(* IEC 61131-3 sources: daoli-st-library/DL_Process (part 52) *)

(* ---- FB_DL_SputterTargetBurnInSeq.st ---- *)
//==============================================================================
// 功能块：FB_DL_SputterTargetBurnInSeq ｜ 中文名称：溅射靶预烧与功率爬坡序（复杂度 C4）
// 所属子库：DL_Process ｜ 版本 VERSION: v1.0.0 ｜ 兼容：CODESYS V3.5+ / TwinCAT 3 / 汇川 InoProShop
// 功能描述：新靶装机后的预烧处理——真空达标 → 通 Ar 稳气 → 功率按斜率爬升 → 预烧到规定
//           能量 → 按斜率降功率 → 关快门 → 关气 → 完成。全程统计打火次数，超限立即把功率
//           指令压到 0 并锁存 xArcTrip；中止与打火停机一律走三段关断序（降功率 → 关快门
//           → 关气），禁单拍全断（会污染靶面）。
// 开源溯源 (Origin)：道莅原创实现（参考 SEMI F47 与磁控溅射靶预烧工艺惯例 分类与参数
//           域，许可证=MIT，借鉴点=「按斜率爬升 + 累计能量达量停烧 + 打火计数联锁」的
//           预烧序）
// 单位表：气压[Pa] / 功率[kW] / 能量[kWh] / 斜率[kW/s] / 打火[次] / 时间[ms]
// 能量离散积分（本件核心积分，换算写清）：
//   fEnergyKWh = Σ (P[kW] × Δt[s]) ÷ 3600 [s/h]；由 W 折算 kW 的 ÷1000 已含在入口量纲
//   上（若上层以 W 给功率，须先 ÷1000 再进本件），Δt 取 DL_SPT_DT_S 假定 10 ms 周期。
// 错误码表（Process 段 0005，故障窗口 3F11~3F19，信息窗口 3F91）：
//   16#0005_3F11 故障级：组态非法（设定压/容差/设定功率/斜率/能量 <= 0 或打火上限 = 0）
//   16#0005_3F12 故障级：实时量入口非有限（腔压 / 功率 NaN 或 Inf）或幅值超上限，拒算
//   16#0005_3F13 故障级：真空未达标超时（tRampTimeout 内气压未进入设定带）
//   16#0005_3F14 故障级：稳气超时（tRampTimeout 内气压未在带内稳住 tGasStabTime）
//   16#0005_3F15 故障级：功率爬坡超时（tRampTimeout 内未爬到设定功率）
//   16#0005_3F16 故障级：预烧超时（tBurnTimeout 内累计能量未达 fBurnEnergyKWh）
//   16#0005_3F17 故障级：打火超限（累计打火 > nArcLimit，功率立即压 0 并锁存 xArcTrip）
//   16#0005_3F18 故障级：关断序超时（降功率/关快门/关气任一段超 tRampTimeout）
//   16#0005_3F19 故障级兜底：状态机落 ELSE 非法态，全输出断
//   16#0005_3F91 信息级：预烧完成（进入 eDone 拍，不置 bError）
//           故障级码全部锁存回放（R187），唯一清除路径 = bReset 上升沿（含打火锁存）。
// 状态机：E_DL_SputterBurnState（八态：eIdle=0 / eVacCheck=10 / eGasStab=20 / eRampUp=30 /
//           eBurnIn=40 / eRampDown=50 / eDone=60 / eFault=99）。三段关断序不占相位，由
//           内部段号 _uDownStage 驱动（0 降功率 / 1 关快门 / 2 关气）。
// 边界行为：① 真空或气压未进带绝不加功率（eRampUp 入口以 _bVacOk 为唯一前提）；② 打火
//           超限属最高优先级：段 5 在功率生成处先判 _bArcTrip 并压 0，不等状态机；③ 三段
//           关断序每段之间留物理动作时间（DL_SPT_SHUTTER_T / DL_SPT_GAS_T），禁单拍全断；
//           ④ 中止与打火停机共用同一关断序，关断后落 eFault 或 eDone 由 _bArcTrip 决定；
//           ⑤ 八态 CASE 每态显式 + ELSE 兜底 → 3F19 全断。
// 语义假设：① nArcCount 为打火探测器累计计数，本件按增量累加并对上游复位做单调化处理；
//           ② 快门开 = xShutterCmd TRUE 表示靶面暴露给基片，预烧期按工艺允许开快门（挡板
//           由上层另控）；③ 腔压判据用绝对偏差带，不含符号方向。
// 依赖纪律：仅 Standard.library（TON / R_TRIG）；零 GVL、零 VAR_EXTERNAL、零物理地址。
// 修订历史：v1.0.0 2026-11-25 R88 首版（无人值守批次 · 复杂件 C4 · 序号 4）
//==============================================================================

(*------------------------------------------------------------------------------
 * 枚举: E_DL_SputterBurnState（归属本功能块，同文件发布，全库唯一定义）
 * 含义: 预烧相位，与段 8 状态机、段 9 输出置位一一对应。
 *-----------------------------------------------------------------------------*)
TYPE E_DL_SputterBurnState :
(
    eIdle     := 0,  // 空闲：等启动沿 / Idle, awaiting the start edge
    eVacCheck := 10, // 真空核对：腔压进入设定带 / Vacuum check against the pressure band
    eGasStab  := 20, // 稳气：通 Ar 并在带内稳住规定时间 / Argon stabilisation inside the band
    eRampUp   := 30, // 功率爬坡：按斜率爬到设定功率 / Power ramp up to the setpoint
    eBurnIn   := 40, // 预烧：累计能量到量前持续 / Burn-in until the energy target is met
    eRampDown := 50, // 降功率与三段关断 / Power ramp down and the three-stage shutdown
    eDone     := 60, // 完成：预烧结束 / Done, burn-in finished
    eFault    := 99  // 故障：组态/超时/打火/非法态 / Fault, configuration, timeout, arcing or illegal state
);
END_TYPE

FUNCTION_BLOCK FB_DL_SputterTargetBurnInSeq
VAR_INPUT
    xEnable       : BOOL;   // 使能，FALSE 期间按中止处理（走三段关断） [—] / Enable, a drop aborts into the shutdown
    xStart        : BOOL;   // 启动请求，上升沿生效 [—] / Start request, rising edge effective
    xAbort        : BOOL;   // 中止请求，任意拍生效（走三段关断） [—] / Abort request, moves into the shutdown
    xReset        : BOOL;   // 故障复位，上升沿清全部锁存（含打火锁存） [—] / Fault reset, clears all latches
    fChamberPressPa : LREAL; // 腔体实际气压 [Pa] / Actual chamber pressure [Pa]
    fPressSetPa   : LREAL;  // 工艺设定气压 [Pa]，须 > 0 / Process pressure setpoint [Pa]
    fPressTolPa   : LREAL;  // 气压允许偏差 [Pa]，须 > 0 / Allowed pressure tolerance [Pa]
    fPowerKW      : LREAL;  // 实际输出功率 [kW] / Actual delivered power [kW]
    fPowerSetKW   : LREAL;  // 预烧设定功率 [kW]，须 > 0 / Burn-in power setpoint [kW]
    fRampKWperS   : LREAL;  // 功率爬坡/降坡斜率 [kW/s]，须 > 0 / Power ramp rate [kW/s]
    fBurnEnergyKWh: LREAL;  // 预烧目标能量 [kWh]，须 > 0 / Burn-in energy target [kWh]
    nArcCount     : UDINT;  // 打火探测器累计计数 [次] / Arc detector accumulated count
    nArcLimit     : UDINT;  // 打火累计上限 [次]，须 > 0 / Accumulated arc ceiling
    tGasStabTime  : TIME;   // 稳气时长 [ms] / Gas stabilisation time [ms]
    tRampTimeout  : TIME;   // 真空/稳气/爬坡/关断超时 [ms] / Vacuum, gas, ramp and shutdown timeout [ms]
    tBurnTimeout  : TIME;   // 预烧最长允许时间 [ms] / Maximum burn-in time [ms]
END_VAR
VAR_OUTPUT
    fPowerCmdKW     : LREAL;  // 功率指令出口 [kW]，0 = 断功率 / Power command outlet [kW], 0 = off
    xArValveCmd     : BOOL;   // 氩气进气阀命令 [—] / Argon inlet valve command
    xShutterCmd     : BOOL;   // 快门命令（TRUE = 开） [—] / Shutter command, TRUE = open
    bRunning        : BOOL;   // 预烧进行中（非空闲非完成非故障） [—] / Burn-in active
    bDone           : BOOL;   // 预烧完成相电平 [—] / Burn-in done, level in the done phase
    bError          : BOOL;   // 故障级标志，仅故障级码置位 [—] / Fault-class flag, fault-level codes only
    nErrCode        : UDINT;  // 错误码，0 = 无错 [—] / Error code, 0 = none
    fEnergyKWh      : LREAL;  // 累计预烧能量 [kWh] / Accumulated burn-in energy [kWh]
    nArcTotal       : UDINT;  // 累计打火次数 [次] / Accumulated arc count
    xArcTrip        : BOOL;   // 打火超限锁存（bReset 清） [—] / Arc trip latch, cleared by bReset
END_VAR
VAR
    _eState         : E_DL_SputterBurnState := E_DL_SputterBurnState.eIdle; // 当前相位 [—] / Current phase
    _bInit          : BOOL := FALSE;  // 首扫标志，取非判定 [—] / First-scan flag, tested negated
    _fPowerCmd      : LREAL;          // 功率指令斜率限幅后的保持量 [kW] / Held command after rate limiting [kW]
    _fEnergyKWh     : LREAL;          // 内部累计能量 [kWh] / Internal accumulated energy [kWh]
    _nArcTotal      : UDINT;          // 内部累计打火次数 [次] / Internal accumulated arc count
    _nArcPrev       : UDINT;          // 上拍打火计数快照 [次] / Previous-scan arc count snapshot
    _bCfgBad        : BOOL;           // 组态非法锁存 / Illegal configuration latch
    _bCfgOk         : BOOL;           // 本拍组态合法（派生量不锁存） [—] / Configuration legal this scan
    _bSigBad        : BOOL;           // 实时量非有限锁存 / Non-finite process value latch
    _bVacOk         : BOOL;           // 气压在设定带内（派生量） [—] / Pressure inside the setpoint band
    _bArcTrip       : BOOL;           // 打火超限锁存 / Arc trip latch
    _bVacTmo        : BOOL;           // 真空超时锁存 / Vacuum timeout latch
    _bGasTmo        : BOOL;           // 稳气超时锁存 / Gas stabilisation timeout latch
    _bRampTmo       : BOOL;           // 爬坡超时锁存 / Ramp timeout latch
    _bBurnTmo       : BOOL;           // 预烧超时锁存 / Burn-in timeout latch
    _bDownTmo       : BOOL;           // 关断序超时锁存 / Shutdown timeout latch
    _bIllegal       : BOOL;           // 非法状态标志 / Illegal state flag
    _bInfoDone      : BOOL;           // 预烧完成信息当拍标志 / Burn-in done info flag of this scan
    _bAbortReq      : BOOL;           // 中止请求合成（xAbort 或失能） [—] / Combined abort request
    _uDownStage     : UINT;           // 关断段号 0=降功率 1=关快门 2=关气 / Shutdown stage 0 power 1 shutter 2 gas
    rtStart         : R_TRIG;         // 启动沿，段 7 无条件刷新 [—] / Start edge, refreshed in segment 7
    rtReset         : R_TRIG;         // 复位沿，段 7 无条件刷新 [—] / Reset edge, refreshed in segment 7
    tonVac          : TON;            // 真空核对超时 [ms] / Vacuum check timeout [ms]
    tonGas          : TON;            // 稳气计时（仅在带内累计） [ms] / Gas stabilisation timer inside the band
    tonGasMax       : TON;            // 稳气最长允许时间 [ms] / Maximum stabilisation time [ms]
    tonRamp         : TON;            // 功率爬坡超时 [ms] / Ramp timeout [ms]
    tonBurn         : TON;            // 预烧最长允许时间 [ms] / Maximum burn-in time [ms]
    tonShutter      : TON;            // 关快门动作让位 [ms] / Shutter travel dwell [ms]
    tonGasClose     : TON;            // 关气动作让位 [ms] / Gas closing dwell [ms]
    tonDownMax      : TON;            // 关断序总超时 [ms] / Total shutdown timeout [ms]
END_VAR
VAR CONSTANT
    DL_EPS           : LREAL := 1.0E-9;      // 浮点容差零点，兼作除法分母下限 / Float epsilon, also the divisor floor
    DL_SPT_DT_S      : LREAL := 0.01;        // 爬坡与积分的假定任务周期 [s]（10 ms） / Assumed task period [s]
    DL_SPT_SEC_PER_H : LREAL := 3600.0;      // 秒折算小时 [s/h]，能量积分用 / Seconds per hour for the energy integral
    DL_SPT_POW_EPS   : LREAL := 0.05;        // 功率到位容差 [kW] / Power arrival tolerance [kW]
    DL_SPT_POWER_MAX : LREAL := 500.0;       // 功率反馈合法幅值上限 [kW] / Legal power ceiling [kW]
    DL_SPT_PRESS_MAX : LREAL := 100000.0;    // 气压反馈合法幅值上限 [Pa] / Legal pressure ceiling [Pa]
    DL_SPT_SHUTTER_T : TIME  := T#800MS;     // 关快门动作让位 [ms] / Shutter travel dwell [ms]
    DL_SPT_GAS_T     : TIME  := T#500MS;     // 关气动作让位 [ms] / Gas closing dwell [ms]
END_VAR
(*------------------------------------------------------------------------------
 * 段 1｜每拍预置：全部输出先落安全侧，单拍标志预清零
 *      All outputs preset to the safe side, one-shot flags pre-cleared
 *-----------------------------------------------------------------------------*)
fPowerCmdKW := 0.0;                         // 功率指令先归零（安全侧） / Power command zeroed first
xArValveCmd := FALSE; xShutterCmd := FALSE; // 氩气与快门命令先断 / Argon and shutter commands cleared
bRunning := FALSE;  bDone := FALSE;         // 运行与完成标志每拍重算 / Running and done flags recomputed
bError := FALSE;    nErrCode := 16#0000_0000; // 故障标志与错误码每拍重算 / Fault flag and code recomputed
_bIllegal := FALSE; _bInfoDone := FALSE;    // 非法态与完成信息预清零 / Illegal and done-info flags pre-cleared

(*------------------------------------------------------------------------------
 * 段 2｜首扫初始化：相位、指令保持量、能量、打火累计与关断段号复位
 *      First-scan initialisation of phase, command, energy, arc count and stage
 *-----------------------------------------------------------------------------*)
IF NOT _bInit THEN
    _eState     := E_DL_SputterBurnState.eIdle; // 相位从空闲起步 / Phase starts idle
    _fPowerCmd := 0.0;  _fEnergyKWh := 0.0;     // 指令与能量从零起步 / Command and energy start at zero
    _nArcTotal := 0;    _nArcPrev  := 0;  _uDownStage := 0; // 打火累计/快照/关断段号从零起步 / Arc, snapshot and stage zero
    _bInit := TRUE;                             // 首扫只做一次 / The first scan runs once
END_IF
(*------------------------------------------------------------------------------
 * 段 3｜实时量入口非有限闸 + 组态闸 + 气压带判据
 *      Non-finite inlet gate, configuration gates and the pressure band criterion
 *-----------------------------------------------------------------------------*)
IF NOT (fChamberPressPa > -1.0E30 AND fChamberPressPa < 1.0E30) THEN _bSigBad := TRUE; END_IF  // 腔压非有限 → 3F12 / Non-finite pressure, 3F12
IF ABS(fChamberPressPa) > DL_SPT_PRESS_MAX THEN _bSigBad := TRUE; END_IF                     // 腔压幅值超上限 → 3F12 / Beyond the ceiling, 3F12
IF NOT (fPowerKW > -1.0E30 AND fPowerKW < 1.0E30) THEN _bSigBad := TRUE; END_IF               // 功率非有限 → 3F12 / Non-finite power, 3F12
IF ABS(fPowerKW) > DL_SPT_POWER_MAX THEN _bSigBad := TRUE; END_IF                             // 功率幅值超上限 → 3F12 / Beyond the ceiling, 3F12
IF NOT (fPressSetPa > -1.0E30 AND fPressSetPa < 1.0E30) THEN _bCfgBad := TRUE; END_IF         // 设定压非有限 → 3F11 / Non-finite setpoint pressure, 3F11
IF NOT (fPowerSetKW > -1.0E30 AND fPowerSetKW < 1.0E30) THEN _bCfgBad := TRUE; END_IF         // 设定功率非有限 → 3F11 / Non-finite setpoint power, 3F11
IF NOT (fRampKWperS > -1.0E30 AND fRampKWperS < 1.0E30) THEN _bCfgBad := TRUE; END_IF         // 斜率非有限 → 3F11 / Non-finite ramp, 3F11
IF NOT (fBurnEnergyKWh > -1.0E30 AND fBurnEnergyKWh < 1.0E30) THEN _bCfgBad := TRUE; END_IF    // 目标能量非有限 → 3F11 / Non-finite energy, 3F11
IF (fPressSetPa <= DL_EPS) OR (fPressTolPa <= DL_EPS) OR (fPowerSetKW <= DL_EPS)
   OR (fRampKWperS <= DL_EPS) OR (fBurnEnergyKWh <= DL_EPS) THEN _bCfgBad := TRUE; END_IF // 五者须为正 → 3F11 / All five must be positive
IF nArcLimit = 0 THEN _bCfgBad := TRUE; END_IF                          // 打火上限为 0 即永久跳闸 → 3F11 / Zero arc limit, 3F11
IF (tGasStabTime <= T#0MS) OR (tRampTimeout <= T#0MS) OR (tBurnTimeout <= T#0MS) THEN _bCfgBad := TRUE; END_IF // 时间量须为正 → 3F11
_bCfgOk := NOT _bCfgBad;                    // 本拍组态合法派生量 / Configuration-legal derived flag of this scan
_bVacOk := ABS(fChamberPressPa - fPressSetPa) <= fPressTolPa; // 气压带判据 [Pa] / Pressure band criterion [Pa]

(*------------------------------------------------------------------------------
 * 段 4｜打火累计（增量单调化）与超限锁存
 *      Arc accumulation with monotonic handling of an upstream counter reset
 *-----------------------------------------------------------------------------*)
IF nArcCount >= _nArcPrev THEN _nArcTotal := _nArcTotal + (nArcCount - _nArcPrev); // 增量累加 / Increment accumulated
ELSE _nArcTotal := _nArcTotal + nArcCount; END_IF                                  // 上游复位按新窗累加 / Upstream reset, new window
_nArcPrev := nArcCount;                     // 计数快照推进 / Count snapshot advanced
IF (_nArcTotal > nArcLimit) THEN
    _bArcTrip := TRUE;                      // 打火超限锁存 → 3F17 / Arc ceiling exceeded, 3F17
END_IF

(*------------------------------------------------------------------------------
 * 段 5｜功率指令生成（打火优先压 0）+ 斜率限幅 + 能量离散积分
 *      Power command generation, arc-first zeroing, rate limiting and energy integral
 *-----------------------------------------------------------------------------*)
IF _bArcTrip THEN
    _fPowerCmd := 0.0;                      // 打火超限：功率立即压 0（不等状态机） / Arc trip, power forced to zero
ELSIF (_eState = E_DL_SputterBurnState.eRampUp) OR (_eState = E_DL_SputterBurnState.eBurnIn) THEN
    IF fPowerSetKW > _fPowerCmd THEN
        _fPowerCmd := _fPowerCmd + fRampKWperS * DL_SPT_DT_S;       // 升坡 [kW] / Ramp up [kW]
        IF _fPowerCmd > fPowerSetKW THEN _fPowerCmd := fPowerSetKW; END_IF // 上钳设定值 / Clamp at setpoint
    ELSIF fPowerSetKW < _fPowerCmd THEN
        _fPowerCmd := _fPowerCmd - fRampKWperS * DL_SPT_DT_S;       // 降坡 [kW] / Ramp down [kW]
        IF _fPowerCmd < fPowerSetKW THEN _fPowerCmd := fPowerSetKW; END_IF // 下钳设定值 / Clamp at setpoint
    END_IF
ELSIF _eState = E_DL_SputterBurnState.eRampDown THEN
    _fPowerCmd := _fPowerCmd - fRampKWperS * DL_SPT_DT_S;           // 关断序段 0：降功率 [kW] / Shutdown stage 0, ramp down
    IF _fPowerCmd < 0.0 THEN _fPowerCmd := 0.0; END_IF              // 下钳 0 / Lower clamp at zero
ELSE
    _fPowerCmd := 0.0;                      // 其余相指令归零 / Zeroed in all other phases
END_IF
IF (_eState = E_DL_SputterBurnState.eBurnIn) AND (DL_SPT_SEC_PER_H > DL_EPS) THEN
    _fEnergyKWh := _fEnergyKWh + (_fPowerCmd * DL_SPT_DT_S) / DL_SPT_SEC_PER_H; // 能量积分 [kWh] / Energy integral [kWh]
END_IF
fPowerCmdKW := _fPowerCmd; fEnergyKWh := _fEnergyKWh; // 功率指令与能量出口 [kW]/[kWh] / Power and energy outlets
nArcTotal := _nArcTotal;    xArcTrip := _bArcTrip;    // 累计打火与打火锁存出口 / Arc count and arc trip outlets

(*------------------------------------------------------------------------------
 * 段 6｜中止入口（任意运行相 → 三段关断序）与复位
 *      Abort entry into the three-stage shutdown plus the reset edge
 *-----------------------------------------------------------------------------*)
_bAbortReq := xAbort OR (NOT xEnable);      // 中止请求合成：显式中止或失能 / Combined abort: explicit abort or enable loss
IF _bAbortReq AND (_eState <> E_DL_SputterBurnState.eIdle) AND (_eState <> E_DL_SputterBurnState.eRampDown)
   AND (_eState <> E_DL_SputterBurnState.eDone) AND (_eState <> E_DL_SputterBurnState.eFault) THEN
    _uDownStage := 0;                       // 关断序从段 0（降功率）起 / Shutdown starts at stage 0
    _eState     := E_DL_SputterBurnState.eRampDown; // 进关断相 / To the shutdown phase
END_IF
IF rtReset.Q THEN
    _bCfgBad := FALSE;  _bSigBad := FALSE;  _bArcTrip := FALSE; // 复位清组态/入口/打火锁存 / Clears configuration, inlet and arc latches
    _bVacTmo := FALSE;  _bGasTmo := FALSE;  _bRampTmo := FALSE; // 复位清真空/稳气/爬坡锁存 / Clears vacuum, gas and ramp latches
    _bBurnTmo := FALSE; _bDownTmo := FALSE;                     // 复位清预烧/关断锁存 / Clears burn-in and shutdown latches
END_IF
(*------------------------------------------------------------------------------
 * 段 7｜定时器与边沿无条件周期刷新（R7：CASE 之外每拍必调，各司其职不复用）
 *      Timers and edges refreshed unconditionally every scan, outside the CASE
 *-----------------------------------------------------------------------------*)
rtStart(CLK := xStart); rtReset(CLK := xReset); // 启动沿与复位沿无条件刷新 / Start and reset edges refreshed
tonVac(IN := (_eState = E_DL_SputterBurnState.eVacCheck), PT := tRampTimeout);                     // 真空核对超时 / Vacuum timeout
tonGas(IN := (_eState = E_DL_SputterBurnState.eGasStab) AND _bVacOk, PT := tGasStabTime);          // 带内稳气计时 / In-band gas timer
tonGasMax(IN := (_eState = E_DL_SputterBurnState.eGasStab), PT := tRampTimeout);                   // 稳气最长允许 / Maximum stabilisation
tonRamp(IN := (_eState = E_DL_SputterBurnState.eRampUp), PT := tRampTimeout);                      // 爬坡超时 / Ramp timeout
tonBurn(IN := (_eState = E_DL_SputterBurnState.eBurnIn), PT := tBurnTimeout);                      // 预烧超时 / Burn-in timeout
tonShutter(IN := (_eState = E_DL_SputterBurnState.eRampDown) AND (_uDownStage = 1), PT := DL_SPT_SHUTTER_T); // 关快门让位 / Shutter dwell
tonGasClose(IN := (_eState = E_DL_SputterBurnState.eRampDown) AND (_uDownStage = 2), PT := DL_SPT_GAS_T);    // 关气让位 / Gas dwell
tonDownMax(IN := (_eState = E_DL_SputterBurnState.eRampDown), PT := tRampTimeout);                  // 关断序总超时 / Shutdown timeout

(*------------------------------------------------------------------------------
 * 段 8｜状态机（含三段关断序；打火停机与中止共用关断序）
 *      Phase machine with the three-stage shutdown shared by abort and arc trip
 *-----------------------------------------------------------------------------*)
CASE _eState OF
    E_DL_SputterBurnState.eIdle:            // 空闲：启动沿 + 组态合法 + 入口可用才进真空核对 / Idle, legal start edge only
        IF rtStart.Q AND _bCfgOk AND (NOT _bSigBad) AND (NOT _bArcTrip) AND (NOT _bAbortReq) THEN
            _fEnergyKWh := 0.0; _nArcTotal := 0; _nArcPrev := nArcCount; // 新靶计数与能量清零 / New target, counters reset
            _uDownStage := 0;               // 关断段号复位 / Shutdown stage reset
            _eState := E_DL_SputterBurnState.eVacCheck; // 进真空核对相 / To the vacuum check
        END_IF
    E_DL_SputterBurnState.eVacCheck:        // 真空核对：气压进带即稳气，超时落故障 / Into the band or time out
        IF _bVacOk THEN _eState := E_DL_SputterBurnState.eGasStab; // 进带，进稳气相 / In band, to stabilisation
        ELSIF tonVac.Q THEN _bVacTmo := TRUE; _eState := E_DL_SputterBurnState.eFault; // 真空超时 → 3F13 / Vacuum timeout, 3F13
        END_IF
    E_DL_SputterBurnState.eGasStab:         // 稳气：带内累计满即爬坡；离带重置；总时超落故障 / In-band accumulation
        IF tonGasMax.Q THEN _bGasTmo := TRUE; _eState := E_DL_SputterBurnState.eFault; // 稳气超时 → 3F14 / Gas timeout, 3F14
        ELSIF tonGas.Q THEN _eState := E_DL_SputterBurnState.eRampUp; // 稳气完成，进爬坡相 / Stabilised, to ramp up
        END_IF
    E_DL_SputterBurnState.eRampUp:          // 爬坡：气压须仍在带内，到设定功率即预烧 / Ramp with the band still proven
        IF NOT _bVacOk THEN _bGasTmo := TRUE; _eState := E_DL_SputterBurnState.eFault; // 爬坡期气压离带 → 3F14 / Band lost, 3F14
        ELSIF _bArcTrip THEN _uDownStage := 0; _eState := E_DL_SputterBurnState.eRampDown; // 打火停机走关断序 / Arc trip, shutdown
        ELSIF ABS(_fPowerCmd - fPowerSetKW) <= DL_SPT_POW_EPS THEN _eState := E_DL_SputterBurnState.eBurnIn; // 到功率，进预烧
        ELSIF tonRamp.Q THEN _bRampTmo := TRUE; _eState := E_DL_SputterBurnState.eFault; // 爬坡超时 → 3F15 / Ramp timeout, 3F15
        END_IF
    E_DL_SputterBurnState.eBurnIn:          // 预烧：能量到量进关断，打火超限立即关断，超时落故障 / Energy or arc or timeout
        IF _bArcTrip THEN _uDownStage := 0; _eState := E_DL_SputterBurnState.eRampDown; // 打火停机走关断序 / Arc trip, shutdown
        ELSIF _fEnergyKWh >= fBurnEnergyKWh THEN _uDownStage := 0; _eState := E_DL_SputterBurnState.eRampDown; // 能量到量，降功率
        ELSIF tonBurn.Q THEN _bBurnTmo := TRUE; _eState := E_DL_SputterBurnState.eFault; // 预烧超时 → 3F16 / Burn-in timeout, 3F16
        END_IF
    E_DL_SputterBurnState.eRampDown:        // 三段关断：0 降功率 → 1 关快门 → 2 关气 → 完成/故障
        IF tonDownMax.Q AND (_uDownStage < 2) THEN _bDownTmo := TRUE; _eState := E_DL_SputterBurnState.eFault; // 关断超时 → 3F18
        ELSIF (_uDownStage = 0) AND (_fPowerCmd <= DL_SPT_POW_EPS) THEN _uDownStage := 1; // 功率到 0，关快门 / Power zero, shutter off
        ELSIF (_uDownStage = 1) AND tonShutter.Q THEN _uDownStage := 2;                   // 快门让位，关气 / Shutter dwelled, gas off
        ELSIF (_uDownStage = 2) AND tonGasClose.Q THEN
            IF _bArcTrip THEN _eState := E_DL_SputterBurnState.eFault;                    // 打火停机落故障 / Arc trip, fault
            ELSE _bInfoDone := TRUE; _eState := E_DL_SputterBurnState.eDone; END_IF         // 正常完成 / Normal completion
        END_IF
    E_DL_SputterBurnState.eDone:            // 完成：启动撤销才回空闲 / Done, back to idle once start drops
        IF NOT xStart THEN _eState := E_DL_SputterBurnState.eIdle; END_IF
    E_DL_SputterBurnState.eFault:           // 故障：复位沿且组态合法且入口可用才回空闲 / Fault, reset edge only
        IF rtReset.Q AND _bCfgOk AND (NOT _bSigBad) THEN _eState := E_DL_SputterBurnState.eIdle; END_IF
    ELSE                                    // 非法状态兜底（R6：CASE 必带 ELSE）/ Illegal-state fallback
        _bIllegal := TRUE; _eState := E_DL_SputterBurnState.eFault; // 非法态 → 3F19，落故障 / Illegal state, 3F19
END_CASE

(*------------------------------------------------------------------------------
 * 段 9｜输出置位（三段关断序：功率→快门→气；打火锁存期严禁再进气或开快门）
 *      Output assignment, the three-stage order, no gas or shutter while tripped
 *-----------------------------------------------------------------------------*)
CASE _eState OF
    E_DL_SputterBurnState.eGasStab:         // 稳气相：只开氩气 / Stabilisation, argon only
        xArValveCmd := TRUE;
    E_DL_SputterBurnState.eRampUp:          // 爬坡相：氩气 + 快门开 / Ramp up with argon and the shutter open
        xArValveCmd := TRUE; xShutterCmd := TRUE;
    E_DL_SputterBurnState.eBurnIn:          // 预烧相：氩气 + 快门开 / Burn-in with argon and the shutter open
        xArValveCmd := TRUE; xShutterCmd := TRUE;
    E_DL_SputterBurnState.eRampDown:        // 关断相：按段号逐级断开 / Shutdown, staged
        xArValveCmd := (_uDownStage < 2);   // 段 2 才关气 / Gas closes at stage 2
        xShutterCmd := (_uDownStage < 1);   // 段 1 才关快门 / Shutter closes at stage 1
    E_DL_SputterBurnState.eDone:            // 完成相：完成电平，两阀全关 / Done, done level and both closed
        bDone := TRUE;
    ELSE                                    // 其余相（空闲/核对/故障）全断 / Other phases, all off
        xArValveCmd := FALSE; xShutterCmd := FALSE;
END_CASE
bRunning := (_eState <> E_DL_SputterBurnState.eIdle) AND (_eState <> E_DL_SputterBurnState.eDone)
            AND (_eState <> E_DL_SputterBurnState.eFault); // 运行标志 / Running flag

(*------------------------------------------------------------------------------
 * 段 10｜错误码映射（锁存回放，R187：故障相不按当下输入重推断）
 *      Error-code map, latched replay
 *-----------------------------------------------------------------------------*)
IF _bIllegal THEN nErrCode := 16#0005_3F19; bError := TRUE;        // 故障级兜底：非法态 / Fault, illegal state fallback
ELSIF _bCfgBad THEN nErrCode := 16#0005_3F11; bError := TRUE;      // 故障级：组态非法 / Fault, illegal configuration
ELSIF _bSigBad THEN nErrCode := 16#0005_3F12; bError := TRUE;      // 故障级：入口非有限 / Fault, non-finite inlet
ELSIF _bArcTrip THEN nErrCode := 16#0005_3F17; bError := TRUE;     // 故障级：打火超限 / Fault, arc trip
ELSIF _bVacTmo THEN nErrCode := 16#0005_3F13; bError := TRUE;      // 故障级：真空超时 / Fault, vacuum timeout
ELSIF _bGasTmo THEN nErrCode := 16#0005_3F14; bError := TRUE;      // 故障级：稳气超时或离带 / Fault, gas timeout or band loss
ELSIF _bRampTmo THEN nErrCode := 16#0005_3F15; bError := TRUE;     // 故障级：爬坡超时 / Fault, ramp timeout
ELSIF _bBurnTmo THEN nErrCode := 16#0005_3F16; bError := TRUE;     // 故障级：预烧超时 / Fault, burn-in timeout
ELSIF _bDownTmo THEN nErrCode := 16#0005_3F18; bError := TRUE;     // 故障级：关断序超时 / Fault, shutdown timeout
ELSIF _bInfoDone THEN nErrCode := 16#0005_3F91;                    // 信息级：预烧完成 / Info, burn-in done
END_IF
END_FUNCTION_BLOCK

(* ---- FB_DL_StackPressureProfile.st ---- *)
(*
  Component : FB_DL_StackPressureProfile
  Category  : DL_Process
  Type      : FB
  Version   : 1.0.0
  CodeSeg   : 16#06_0_39
  Summary   : 叠片压力曲线与保压判定：压力段轮廓（升压-保压-泄压）+ 保压容差窗 + 越窗分级。
              Stacking pressure profile and hold verdict: ramp-hold-release segments with a tolerance window and graded verdict.
  溯源声明  : 参照 FB_DL_RampSoakProfile 段轮廓骨架语义，clean-room 自含实现，无实例依赖
  边界安全  : 压力非有限（NaN 自反 + Inf 上限）与负值域拦截；段时长正域闸（> 0，防状态机卡死）；
              容差域闸（> 0）；段进度按节拍计数（自复位 TON），越过段尾推进；压力单位 kN 全程标注；
              保压窗判定带容差比较（禁等值直比）；判定结果锁存至下一周期起动沿解除（可达路径）。
  复用      : 参照 FB_DL_RampSoakProfile 骨架语义（clean-room 自含实现，无实例依赖）
*)

FUNCTION_BLOCK FB_DL_StackPressureProfile
VAR_INPUT
    bRun      : BOOL;                   (* 周期使能/起动 [事件] · Cycle enable/start *)
    fPressKN  : LREAL;                  (* 实测压力 [kN] · Measured pressure *)
    fRampKN   : LREAL := 12.0;          (* 升压段目标 [kN] · Ramp target *)
    fHoldKN   : LREAL := 10.0;          (* 保压段目标 [kN] · Hold target *)
    tRampMs   : TIME  := T#2000MS;      (* 升压段时长 [ms] · Ramp duration *)
    tHoldMs   : TIME  := T#3000MS;      (* 保压段时长 [ms] · Hold duration *)
    fTolKN    : LREAL := 0.5;           (* 保压容差 [kN] · Hold tolerance *)
    fEps      : LREAL := 1.0E-6;        (* 浮点判零容差 [实数域] · Floating zero tolerance *)
END_VAR
VAR_OUTPUT
    ePhase  : (ePhIdle := 0, ePhRamp := 1, ePhHold := 2, ePhRelease := 3);  (* 相枚举输出 / Phase output enum *)
    fTargetKN: LREAL;                   (* 当前段目标压力 [kN] · Current segment target *)
    bInWin  : BOOL;                     (* 本拍在保压容差窗内 [开关] · In the hold window *)
    nViolN  : INT;                      (* 本周期越窗拍数 [拍] · Violation scans this cycle *)
    bError  : BOOL;                     (* 故障标志，与故障码配对 · Fault flag paired with codes *)
    uErrorId: UDINT;                    (* 事件码 16#0000_0039，0 无事件 · Event code *)
END_VAR
VAR
    _eState : (eStIdle := 0, eStRamp := 1, eStHold := 2, eStRelease := 3);  (* 内部状态机 / Internal state machine *)
    uCode   : WORD;     (* 码位暂存，每拍重算 [码] · Code staging *)
    tonSeg  : TON;      (* 段计时 [ms]，自复位振荡 · Segment timer, self-reset *)
    bSigOk  : BOOL;     (* 输入有效标志 · Input validity flag *)
    bRunPrv : BOOL;     (* 上拍起动快照，上升沿判据 · Previous run snapshot *)
    bStart  : BOOL;     (* 起动上升沿 [脉冲] · Start rising edge *)
    nCycles : UDINT;    (* 完成周期计数 [次]，防回卷 · Completed cycle count *)
END_VAR
VAR CONSTANT
    DL_SPP_WRAP : UDINT := 4294967290;  (* 计数防回卷余量 [次] · Counter wrap guard *)
END_VAR

(* === 段 0 · 实例刷新（每拍无条件，红线 7）=== *)
tonSeg(IN := NOT tonSeg.Q, PT := T#100MS);      (* 段进度节拍自复位振荡 / Self-reset progress pace *)
bStart := bRun AND (NOT bRunPrv);               (* 起动上升沿 / Start edge *)
bRunPrv := bRun;                                (* 快照更新 / Snapshot *)

(* === 段 1 · 输入校验与量程闸 === *)
uCode := 16#0000;                       // 每拍清码（可达清零基线）/ Clear codes each scan
bSigOk := (fPressKN = fPressKN) AND (ABS(fPressKN) < 1.0E308)   // 非有限拦截 / Non-finite guard
          AND (fPressKN >= 0.0)                                          // 压力非负域闸 / Non-negative pressure
          AND (fTolKN > fEps)                                            // 容差正域闸 / Tolerance gate
          AND (tRampMs > T#0MS) AND (tHoldMs > T#0MS);                   // 段时长正域闸 / Duration gates
IF NOT bSigOk THEN
    uCode := 16#0039;                   // 故障级：域外，轮廓冻结 / Fault: domain invalid
END_IF

(* === 段 2 · 主逻辑：三段轮廓状态机 === *)
IF bStart AND bSigOk THEN
    _eState := eStRamp;                 (* 拍 N 起动沿进入，拍 N+1 升压相 / To ramp on start edge *)
    nViolN := 0;                        (* 新周期越窗计数清零 / Reset violation count *)
    tonSeg(IN := FALSE, PT := T#100MS); (* 段计时复位重启 / Restart the segment timer *)
END_IF
IF bSigOk THEN
    CASE _eState OF
        eStIdle:                        (* 空闲相：目标钳零 / Idle: zero target *)
            fTargetKN := 0.0;           (* 目标零压 / Zero target *)
        eStRamp:                        (* 升压相：目标=升压目标；窗满转保压 / Ramp *)
            fTargetKN := fRampKN;       (* 升压目标 [kN] / Ramp target *)
            IF tonSeg.Q OR (fPressKN >= (fRampKN - fEps)) THEN
                _eState := eStHold;     (* 时窗满或到位转保压 / To hold on time or arrival *)
                tonSeg(IN := FALSE, PT := tHoldMs);     (* 重载保压时长 / Reload hold duration *)
            END_IF
        eStHold:                        (* 保压相：容差窗判定与越窗计数 / Hold: tolerance verdict *)
            fTargetKN := fHoldKN;       (* 保压目标 [kN] / Hold target *)
            bInWin := (fPressKN > (fHoldKN - fTolKN)) AND (fPressKN < (fHoldKN + fTolKN));
                                        (* 容差窗判定（带限非等比）/ In-window verdict *)
            IF NOT bInWin THEN
                nViolN := nViolN + 1;   (* 越窗拍累加 / Count violations *)
            END_IF
            IF tonSeg.Q THEN
                _eState := eStRelease;  (* 保压窗满转泄压 / To release *)
                tonSeg(IN := FALSE, PT := T#100MS);
            END_IF
        eStRelease:                     (* 泄压相：目标回零，到位收周期 / Release *)
            fTargetKN := 0.0;           (* 泄压目标零 [kN] / Release to zero *)
            IF fPressKN < fEps THEN
                _eState := eStIdle;     (* 到位回空闲，周期收口 / Back to idle *)
                IF nCycles < DL_SPP_WRAP THEN
                    nCycles := nCycles + 1;     (* 完成周期计数 / Count the cycle *)
                END_IF
            END_IF
    ELSE
        _eState := eStIdle;             (* ELSE 兜底回空闲安全相 / ELSE fallback to idle *)
        fTargetKN := 0.0;
        uCode := 16#0039;               (* 状态越界报码 / Code on illegal state *)
    END_CASE
END_IF

(* === 段 3 · 输出映射与故障码（CASE 内未触碰输出枚举）=== *)
ePhase := ePhIdle;                      (* 相映射默认 / Default mapping *)
IF _eState = eStRamp THEN
    ePhase := ePhRamp;                  (* 升压相映射 / Map ramp *)
ELSIF _eState = eStHold THEN
    ePhase := ePhHold;                  (* 保压相映射 / Map hold *)
ELSIF _eState = eStRelease THEN
    ePhase := ePhRelease;               (* 泄压相映射 / Map release *)
END_IF
IF _eState <> eStHold THEN
    bInWin := FALSE;                    (* 非保压相在窗标志清零 / Clear in-window outside hold *)
END_IF
bError := (uCode <> 16#0000);           (* 故障标志配对 / Fault flag paired *)
uErrorId := WORD_TO_UDINT(uCode);       (* 码位单点写入（16#0000_0039 形态）/ Single write point *)
END_FUNCTION_BLOCK

(* ---- FB_DL_StakingPressCtrl.st ---- *)
(*
  FB_DL_StakingPressCtrl  —  叠片台压装顺控（对齐-压紧-保压-泄压 + 压力窗判据） / Stacking-table press-fit sequencer with pressure-window verdict
  分类 Category : DL_Process
  版本 Version  : 1.0.0
  来源 Source   : roadmap-li-p1 — 锂电叠片工站压装顺控真缺口
  溯源 Origin   : 道莅 clean-room 实现；压装四段（对齐/压紧/保压/泄压）时序与压力窗判据为公开工艺逻辑，未复制任何源码行
  功能 Function : 1) 四段顺控：eAlign 对齐（等 bAlignInPos 且 tAlign 到时）→ ePress 压紧
                  （等 fPressMpa >= fWinLoMpa）→ eHold 保压（tHold 计时，窗内保持）→
                  eVent 泄压（tVent 计时）→ eDone；2) 压力窗判据：保压相 fPressMpa 越
                  [fWinLoMpa, fWinHiMpa] 即故障；3) 超时保护：对齐/压紧/泄压三相各有独立
                  TON，超时即故障；4) 故障级单码 039D，归因由 eCause 独立枚举成员承载
                  （组态非法/对齐超时/压紧超时/保压越窗/泄压超时，R190 归因唯一）；
                  5) 信息级 04C5 = 压装循环完成沿；6) 解除式全当拍量（R240）。
  接口 Interface: 输入 8 个工艺量 + 4 个时间量 + 3 个命令位；输出状态/压力镜像/原因/故障码
  边界 Boundary : ① 组态闸：fWinLoMpa < 0.0、fWinHiMpa <= fWinLoMpa、四个时间量 <= T#0S
                  任一成立 → 039D 锁存且 eCause = eCfgIllegal；
                  ② 浮点比较全部容差式（ABS 差值 < 1.0E-6），禁 = / <> 判等；
                  ③ 四个 TON 实例均在段 0 无条件每周期调用，IN 由相位判据派生，相切换
                  自动复位 ET，无跨相残留（R176）；
                  ④ 故障相迁出唯一路径 = bReset 上升沿（段 4 承载），禁死锁；
                  ⑤ 零全局耦合：无 GVL / VAR_EXTERNAL / %I %Q %M 直接地址。
  依赖 Depends  : Standard.library（TON / R_TRIG）
  码表 Error codes（Process 段 0005，故障窗口 039D / 信息窗口 04C5）:
    16#0005_039D 故障级：压装故障总码（组态非法 / 对齐超时 / 压紧超时 / 保压越窗 / 泄压超时），
                 锁存至 bReset 上升沿；逐成因归因见 eCause，不新增码位（派单硬约束单码）
    16#0005_04C5 信息级：压装循环完成沿（泄压完成进 eDone 单拍）
  修订历史 Revision :
    2026-11-19  v1.0.0  R43 首版（批次 1 · 序号 1）
*)

TYPE E_DL_SpcState :
(
    eIdle   := 0,     // 未使能待启动 / Idle, waiting for start
    eAlign  := 10,    // 对齐中，等对位信号 / Aligning, waiting alignment
    ePress  := 20,    // 压紧中，等压力达窗下限 / Pressing, waiting pressure reaching window
    eHold   := 30,    // 保压中，计时并在窗内保持 / Holding with window supervision
    eVent   := 40,    // 泄压中，等泄压到时 / Venting, waiting vent time
    eDone   := 50,    // 循环完成，待撤启动 / Done, waiting start release
    eFault  := 90     // 故障锁存相 / Fault latched phase
);
END_TYPE

TYPE E_DL_SpcCause :
(
    eNone        := 0,    // 无故障成因 / No cause
    eCfgIllegal  := 1,    // 组态非法（窗口/时间域非法） / Illegal configuration
    eAlignTmo    := 2,    // 对齐超时 / Alignment timeout
    ePressTmo    := 3,    // 压紧超时（未达窗下限） / Press timeout
    eHoldDev     := 4,    // 保压越窗 / Hold pressure out of window
    eVentTmo     := 5     // 泄压超时 / Vent timeout
);
END_TYPE

FUNCTION_BLOCK FB_DL_StakingPressCtrl
VAR_INPUT
    fPressMpa    : REAL := 0.0;        // 实测压装压力 [MPa] / Measured press force
    fWinLoMpa    : REAL := 2.0;        // 压力窗下限 [MPa]，域 >= 0 / Pressure window low limit
    fWinHiMpa    : REAL := 6.0;        // 压力窗上限 [MPa]，域 > 下限 / Pressure window high limit
    tAlign       : TIME := T#2S;       // 对齐超时 [ms]，域 > 0 / Alignment timeout
    tPress       : TIME := T#3S;       // 压紧超时 [ms]，域 > 0 / Press timeout
    tHold        : TIME := T#5S;       // 保压时长 [ms]，域 > 0 / Hold duration
    tVent        : TIME := T#1S;       // 泄压时长 [ms]，域 > 0 / Vent duration
    bAlignInPos  : BOOL := FALSE;      // 对位到位信号（电平）[-] / Alignment-in-position
    bStart       : BOOL := FALSE;      // 启动命令（电平）[-] / Start command, level
    bReset       : BOOL := FALSE;      // 复位命令，上升沿清故障 [-] / Reset edge
END_VAR
VAR_OUTPUT
    eState       : E_DL_SpcState;      // 状态出口，段 6 单点映射 / State outlet
    eCause       : E_DL_SpcCause;      // 故障成因出口（R190 归因唯一） / Fault cause outlet
    fPressMpaOut : REAL;               // 压力镜像 [MPa] / Pressure mirror
    bInWindow    : BOOL;               // 压力在窗内镜像 [-] / Pressure-in-window mirror
    bCycleDone   : BOOL;               // 循环完成标志（eDone 电平）[-] / Cycle done flag
    bError       : BOOL;               // 故障锁存标志 [-] / Fault latch flag
    nErrId       : UDINT;              // 事件码，0 = 无事件 / Event code
END_VAR
VAR
    _eState      : E_DL_SpcState := E_DL_SpcState.eIdle;   // 内部相位（CASE 唯一写入目标） / Internal phase
    _eCause      : E_DL_SpcCause := E_DL_SpcCause.eNone;   // 故障成因锁存（锁存量） / Latched cause
    tonAlign     : TON;                // 对齐计时实例，每周期无条件调用 / Align timer
    tonPress     : TON;                // 压紧计时实例，每周期无条件调用 / Press timer
    tonHold      : TON;                // 保压计时实例，每周期无条件调用 / Hold timer
    tonVent      : TON;                // 泄压计时实例，每周期无条件调用 / Vent timer
    rtReset      : R_TRIG;             // 复位沿实例，每周期无条件调用 / Reset edge
    _bWinOk      : BOOL;               // 压力在窗内当拍量 [-] / Pressure in window, current scan
    _bCfgBad     : BOOL;               // 组态非法当拍量 [-] / Illegal configuration, current scan
    _bFault      : BOOL;               // 故障锁存位（锁存量） / Latched fault bit
    _uFault      : UDINT;              // 故障码锁存（锁存量） / Latched fault code
    _uInfo       : UDINT;              // 信息码，每拍重算 / Transient info code
END_VAR

(* —— 段 0：沿实例与定时器无条件周期刷新（禁置于 IF/CASE 内，IN 由相位判据派生） —— *)
_bWinOk := (fPressMpa >= fWinLoMpa - 1.0E-6) AND (fPressMpa <= fWinHiMpa + 1.0E-6);  // 压力窗判据（容差式） / Window verdict with tolerance
_bCfgBad := (fWinLoMpa < 0.0) OR (fWinHiMpa <= fWinLoMpa)
            OR (tAlign <= T#0S) OR (tPress <= T#0S) OR (tHold <= T#0S) OR (tVent <= T#0S);  // 组态非法当拍量 / Config-illegal current scan
rtReset(CLK := bReset);                                   // 复位沿，每拍必调 / Reset edge refresh
tonAlign(IN := (_eState = E_DL_SpcState.eAlign), PT := tAlign);   // 对齐计时，相外自动复位 ET / Align timer, ET reset out of phase
tonPress(IN := (_eState = E_DL_SpcState.ePress), PT := tPress);   // 压紧计时，相外自动复位 ET / Press timer
tonHold(IN := (_eState = E_DL_SpcState.eHold), PT := tHold);      // 保压计时，相外自动复位 ET / Hold timer
tonVent(IN := (_eState = E_DL_SpcState.eVent), PT := tVent);      // 泄压计时，相外自动复位 ET / Vent timer

(* —— 段 1：单拍量预清零（锁存量 _bFault/_uFault/_eCause 不入清单，禁同拍抹除 R187） —— *)
_uInfo := 16#0000_0000;            // 信息码每拍重算 / Info code recomputed per scan
fPressMpaOut := 0.0;               // 压力镜像缺省 0 / Pressure mirror default
bInWindow := FALSE;                // 窗内镜像缺省 FALSE / Window mirror default
bCycleDone := FALSE;               // 完成标志缺省 FALSE / Done flag default
nErrId := 16#0000_0000;            // 事件码缺省无事件 / Event code default

(* —— 段 2：复位沿 + 组态域闸（当拍量判据） —— *)
IF rtReset.Q THEN                              // rtReset.Q = 当拍量 / current scan
    _bFault := FALSE;                          // 清故障锁存位（锁存量） / Clear fault latch
    _uFault := 16#0000_0000;                   // 清故障锁存码（锁存量） / Clear fault code
    _eCause := E_DL_SpcCause.eNone;            // 清故障成因（锁存量） / Clear cause
    IF _eState = E_DL_SpcState.eFault THEN
        _eState := E_DL_SpcState.eIdle;        // 故障相迁出：回未使能 / Fault exit to idle
    END_IF
END_IF
IF _bCfgBad THEN                               // 组态域闸（当拍量） / Config gate, current scan
    _uFault := 16#0005_039D;                   // 故障级：压装故障总码 / Process fault code
    _eCause := E_DL_SpcCause.eCfgIllegal;      // 归因：组态非法 / Cause: illegal config
    _bFault := TRUE;                           // 故障标志与码位配对（R45） / Flag paired with code
END_IF

(* —— 段 3：分相超时与越窗锁存（判据当拍量；锁存后不再重算成因，故障码锁存回放） —— *)
IF (NOT _bFault) AND tonAlign.Q THEN           // 对齐超时（tonXxx.Q 当拍量） / Align timeout
    _uFault := 16#0005_039D;                   // 故障级：压装故障总码 / Same public code
    _eCause := E_DL_SpcCause.eAlignTmo;        // 归因：对齐超时 / Cause: align timeout
    _bFault := TRUE;
END_IF
IF (NOT _bFault) AND tonPress.Q THEN           // 压紧超时（未达窗下限） / Press timeout
    _uFault := 16#0005_039D;
    _eCause := E_DL_SpcCause.ePressTmo;        // 归因：压紧超时 / Cause: press timeout
    _bFault := TRUE;
END_IF
IF (NOT _bFault) AND (_eState = E_DL_SpcState.eHold) AND (NOT _bWinOk) THEN   // 保压越窗 / Hold out of window
    _uFault := 16#0005_039D;
    _eCause := E_DL_SpcCause.eHoldDev;         // 归因：保压越窗 / Cause: hold deviation
    _bFault := TRUE;
END_IF
IF (NOT _bFault) AND tonVent.Q THEN            // 泄压超时 / Vent timeout
    _uFault := 16#0005_039D;
    _eCause := E_DL_SpcCause.eVentTmo;         // 归因：泄压超时 / Cause: vent timeout
    _bFault := TRUE;
END_IF

(* —— 段 4：故障解除式（R240；全当拍量，逐 BOOL 标注）：
     rtReset.Q = 当拍量；NOT tonAlign.Q / NOT tonPress.Q / NOT tonVent.Q = 当拍量；
     NOT _bCfgBad = 当拍量。组态非法者需先修参数再复位，复位沿当拍组态已合法方可解。 —— *)
IF rtReset.Q AND (NOT _bCfgBad) AND (NOT tonAlign.Q) AND (NOT tonPress.Q) AND (NOT tonVent.Q) THEN
    _bFault := FALSE;                          // 清故障锁存位（锁存量） / Clear fault latch
    _uFault := 16#0000_0000;                   // 清故障锁存码（锁存量） / Clear fault code
    _eCause := E_DL_SpcCause.eNone;            // 清故障成因（锁存量） / Clear cause
END_IF

(* —— 段 4A：故障锁存相位迁移闸（置位后强制入故障相，冻结段 5 内一切推进） —— *)
IF _bFault AND (_eState <> E_DL_SpcState.eFault) THEN
    _eState := E_DL_SpcState.eFault;           // 锁存即入故障相 / Latch enters fault phase
END_IF

(* —— 段 5：相位机（CASE 全覆盖 + ELSE 兜底） —— *)
CASE _eState OF

E_DL_SpcState.eIdle:
    IF bStart AND (NOT _bFault) THEN           // 启动沿条件（电平门 + 无故障） / Start gate
        _eState := E_DL_SpcState.eAlign;       // 进对齐相 / Enter align
    END_IF

E_DL_SpcState.eAlign:
    IF bAlignInPos THEN                        // 出口 1：对位到位（事件量） / Alignment reached
        _eState := E_DL_SpcState.ePress;       // 进压紧相 / Enter press
    ELSIF NOT bStart THEN                      // 出口 2：撤启动（前置消失，R98 双出口） / Start released
        _eState := E_DL_SpcState.eIdle;        // 回未使能 / Back to idle
    END_IF

E_DL_SpcState.ePress:
    IF fPressMpa >= (fWinLoMpa - 1.0E-6) THEN  // 压力达窗下限（容差式） / Pressure reached low limit
        _eState := E_DL_SpcState.eHold;        // 进保压相 / Enter hold
    ELSIF NOT bStart THEN                      // 撤启动：中止本次压装 / Abort on start release
        _eState := E_DL_SpcState.eIdle;
    END_IF

E_DL_SpcState.eHold:
    IF tonHold.Q THEN                          // 保压到时 / Hold elapsed
        _eState := E_DL_SpcState.eVent;        // 进泄压相 / Enter vent
    ELSIF NOT bStart THEN                      // 撤启动：中止 / Abort on start release
        _eState := E_DL_SpcState.eIdle;
    END_IF

E_DL_SpcState.eVent:
    IF tonVent.Q THEN                          // 泄压到时 / Vent elapsed
        _uInfo := 16#0005_04C5;                // 信息级：循环完成沿 / Info: cycle complete edge
        _eState := E_DL_SpcState.eDone;        // 进完成相 / Enter done
    ELSIF NOT bStart THEN                      // 撤启动：中止 / Abort on start release
        _eState := E_DL_SpcState.eIdle;
    END_IF

E_DL_SpcState.eDone:
    IF NOT bStart THEN                         // 撤启动后回空闲（等下一循环） / Start released returns idle
        _eState := E_DL_SpcState.eIdle;
    END_IF

E_DL_SpcState.eFault:
    ;                                          // 故障相：仅段 4 复位沿可迁出 / Fault: only reset edge exits

ELSE
    _uFault := 16#0005_039D;                   // 故障级：非法相位兜底（归并总码，码表声明） / Illegal phase fallback
    _eCause := E_DL_SpcCause.eCfgIllegal;      // 归因：相位非法归并组态 / Cause: phase illegal
    _bFault := TRUE;
    _eState := E_DL_SpcState.eFault;           // 强制回故障相 / Force fault phase

END_CASE

(* —— 段 6：出口单点映射（名实同源；锁存码回放，禁同拍抹除） —— *)
fPressMpaOut := fPressMpa;                     // 压力镜像（名实同源） / Pressure mirror
bInWindow := _bWinOk AND (NOT _bFault);        // 窗内镜像（故障相强制 FALSE） / Window mirror
bCycleDone := (_eState = E_DL_SpcState.eDone); // 完成标志（相电平） / Done flag
IF _bFault THEN
    nErrId := _uFault;                         // 故障锁存码回放 / Replay latched code
ELSE
    nErrId := _uInfo;                          // 信息码（单拍） / Transient info code
END_IF
bError := _bFault;                             // 故障标志与锁存位同源 / Flag from latch
eState := _eState;                             // 状态出口单点映射 / State outlet
eCause := _eCause;                             // 成因出口单点映射 / Cause outlet

END_FUNCTION_BLOCK

(* ---- FB_DL_SteamCondensatePot.st ---- *)
//==============================================================================
// 功能块：FB_DL_SteamCondensatePot ｜ 中文名称：凝液罐液位-排放顺控
// 所属子库：DL_Process ｜ 版本：v1.0.0 ｜ 兼容：CODESYS V3.5+ / TwinCAT 3 / 汇川 InoProShop
// 功能描述：凝液罐液位双限排放顺控——液位达排放启位开排水阀、降至停位
//           关阀（迟滞对），单次排放限时保护（超时液位未降判排放堵塞），
//           排放计数累计。
// 开源溯源 (Origin)：道莅原创实现（参考蒸汽凝液回收系统工程惯例 分类与参数域）
// 单位表：液位[%] / 阈值[%] / 时间[ms] / 计数[次]
// 错误码表：16#0005_01E8 信息级（液位域外已钳位 0~100，不置 bError）/
//           16#0005_01E9 预留禁用（不得挪用）/ 16#0005_0321 故障级（迟滞
//           倒置：停位 >= 启位，组态非法，置 bError）/ 16#0005_0322 故障级
//           （排放超时液位未降，判排放堵塞，关阀，置 bError）/
//           16#0005_0323 故障级兜底（状态机落 ELSE，置 bError）
// 状态机：E_DL_CondPotState（五态：eIdle=0 / eDraining=10 / eTimeout=20 /
//           eReady=30 / eFault=99），CASE 含 ELSE 兜底，ELSE 置 0323 并关阀
// 边界行为：① fPumpLevelLoPct >= fPumpLevelHiPct → 故障 0321（迟滞倒置）；
//           ② 排放超 tDrainMax 液位未降 → 故障 0322 + 关阀（转 eTimeout，
//           bReset 或液位回落解除）；③ 液位域外钳 0~100 + 信息 01E8；
//           ④ 排放计数饱和 4294967295 不回绕；⑤ 液位非有限 → 故障 0321
//           复用（R90，安全侧关阀）。
// 依赖纪律：仅 Standard.library；零跨层调用。
// 修订历史：v1.0.0 2026-11-17 首版（R23 派单 · ROADMAP 公用工程 P1 §392）
//==============================================================================

(*------------------------------------------------------------------------------
 * 枚举: E_DL_CondPotState（归属本功能块，同文件发布，全库唯一定义）
 * 含义: 凝液罐排放相位，每个成员在 CASE 中有且仅有一个标签。
 *-----------------------------------------------------------------------------*)
TYPE E_DL_CondPotState :
(
    eIdle     := 0,   // 空闲：等使能 / Idle, awaiting enable
    eReady    := 10,  // 就绪：液位低于启位，等排放条件 / Ready, level below the start threshold
    eDraining := 20,  // 排放中：排水阀开，等液位降至停位 / Draining, valve open, waiting for the stop level
    eTimeout  := 30,  // 排放超时：判堵塞，阀已关，等解除 / Drain timeout, clog suspected, valve closed
    eFault    := 99   // 故障：组态非法/非有限/非法状态 / Fault, illegal config, non-finite or illegal state
);
END_TYPE

FUNCTION_BLOCK FB_DL_SteamCondensatePot
VAR_INPUT
    fLevelPct        : LREAL;             // 液位实测 [百分数]，有效域 0..100，域外钳位 / Measured level [percent], 0..100, clamped outside
    fPumpLevelHiPct  : LREAL := 80.0;     // 排放启位液位 [百分数] / Drain-start level [percent]
    fPumpLevelLoPct  : LREAL := 30.0;     // 排放停位液位 [百分数]，须 < 启位 / Drain-stop level [percent], must be below the start
    bDrainValveFb    : BOOL;              // 排水阀开反馈 [—] / Drain valve open feedback
    tDrainMax        : TIME  := T#30S;    // 单次排放上限 [ms] / Single-drain ceiling [ms]
    bEnable          : BOOL;              // 使能 [—] / Enable
    bReset           : BOOL;              // 故障复位 [—]，清除超时态 / Fault reset, clears the timeout state
END_VAR
VAR_OUTPUT
    bDrainOut        : BOOL;              // 排水阀输出 [—] / Drain valve output
    ePotState        : E_DL_CondPotState; // 排放相位 [—] / Drain phase
    uDrainCount      : UDINT;             // 排放计数 [次]，饱和不回绕 / Drain counter [count], saturated without wrap
    eErr             : UDINT;             // 错误码，0 = 无错 / Error code, 0 = no error
    bError           : BOOL;              // 故障级标志，仅故障级错误置位 / Fault-class flag, set only on fault-level codes
    bValid           : BOOL;              // 输出可用标志 / Outputs usable flag
END_VAR
VAR
    fbDrainMax       : TON;               // 单次排放限时计时，段 6 无条件刷新 [ms] / Single-drain timer
    _eState          : E_DL_CondPotState := E_DL_CondPotState.eIdle; // 当前相位 / Current phase
    _fLevelEff       : LREAL;             // 钳位后的生效液位 [百分数] / Effective clamped level [percent]
    _bInit           : BOOL := FALSE;     // 首扫标志，初值 FALSE 取非判定 / First-scan flag, tested negated
    _bHystBad        : BOOL;              // 迟滞倒置/非有限锁存 / Hysteresis inversion or non-finite latch
    _bLevelInfo      : BOOL;              // 液位钳位信息当拍标志 / Level clamp info flag of this scan
    _bIllegal        : BOOL;              // 非法状态标志 / Illegal state flag
END_VAR
VAR CONSTANT
    DL_POT_INF       : LREAL := 1.7976931348623157E308; // LREAL 幅值上限 / LREAL magnitude ceiling
    DL_POT_LVL_MIN   : LREAL := 0.0;      // 液位钳位下限 [百分数] / Level clamp floor [percent]
    DL_POT_LVL_MAX   : LREAL := 100.0;    // 液位钳位上限 [百分数] / Level clamp ceiling [percent]
    DL_POT_CNT_MAX   : UDINT := 4294967295; // 排放计数饱和上限 [次] / Drain counter saturation ceiling [count]
END_VAR

(*------------------------------------------------------------------------------
 * 段 1｜每拍预置：阀输出先断（安全侧），单拍标志预清零
 *      Valve output cleared first, fail-safe, one-shot flags pre-cleared
 *-----------------------------------------------------------------------------*)
bDrainOut := FALSE;                         // 排水阀输出先清（安全侧） / Drain output cleared first
eErr      := 16#0000_0000;                  // 错误码每拍重算 / Error code recomputed
bError    := FALSE;                         // 故障标志每拍重算 / Fault flag recomputed
bValid    := FALSE;                         // 可用标志每拍重算 / Usable flag recomputed
_bIllegal := FALSE;                         // 非法状态标志预清零 / Illegal flag pre-cleared
_bLevelInfo := FALSE;                       // 钳位信息预清零 / Clamp info pre-cleared

(*------------------------------------------------------------------------------
 * 段 2｜首扫初始化
 *      First-scan initialisation
 *-----------------------------------------------------------------------------*)
IF NOT _bInit THEN
    _eState   := E_DL_CondPotState.eIdle;   // 相位空闲起步 / Phase starts idle
    uDrainCount := 0;                       // 计数清零 / Counter cleared
    _bHystBad := FALSE;                     // 迟滞锁存清零 / Hysteresis latch cleared
    _bInit    := TRUE;                      // 首扫只做一次 / The first scan runs once
END_IF

(*------------------------------------------------------------------------------
 * 段 3｜组态与输入防御闸（迟滞倒置 / 非有限液位 → 0321 复用，R90）
 *      Configuration and input defense gates, code reused per R90
 *-----------------------------------------------------------------------------*)
IF (fLevelPct <> fLevelPct) OR (ABS(fLevelPct) > DL_POT_INF)
   OR (fPumpLevelHiPct <> fPumpLevelHiPct) OR (ABS(fPumpLevelHiPct) > DL_POT_INF)
   OR (fPumpLevelLoPct <> fPumpLevelLoPct) OR (ABS(fPumpLevelLoPct) > DL_POT_INF) THEN
    _bHystBad := TRUE;                      // 非有限液位/阈值归入迟滞倒置（R90 复用） / Non-finite folded into the inversion fault
END_IF
IF (NOT _bHystBad) AND (fPumpLevelLoPct >= fPumpLevelHiPct) THEN
    _bHystBad := TRUE;                      // 迟滞倒置锁存 / Hysteresis inversion latched
END_IF

(*------------------------------------------------------------------------------
 * 段 4｜液位钳位（域外信息级照算）
 *      Level clamping with an info notice
 *-----------------------------------------------------------------------------*)
IF (NOT _bHystBad) AND ((fLevelPct < DL_POT_LVL_MIN) OR (fLevelPct > DL_POT_LVL_MAX)) THEN
    _fLevelEff := MIN(MAX(fLevelPct, DL_POT_LVL_MIN), DL_POT_LVL_MAX); // 双侧钳位到 0~100 / Two-sided clamp into 0..100
    _bLevelInfo := TRUE;                    // 钳位信息置位 / Clamp info raised
ELSE
    _fLevelEff := fLevelPct;                // 合法液位原值生效 / Valid level applied as-is
END_IF

(*------------------------------------------------------------------------------
 * 段 5｜排放限时计时无条件刷新（R40：CASE 之外每拍必调）
 *      Drain timer refreshed unconditionally per R40
 *-----------------------------------------------------------------------------*)
fbDrainMax(IN := (_eState = E_DL_CondPotState.eDraining) AND bDrainValveFb, PT := tDrainMax); // 排放限时 / Single-drain timer

(*------------------------------------------------------------------------------
 * 段 6｜相位机（只做迁移；输出在段 7 按相置位）
 *      Phase machine, transitions only, outputs assigned in segment seven
 *-----------------------------------------------------------------------------*)
IF _bHystBad THEN
    _eState := E_DL_CondPotState.eFault;    // 组态/输入异常直接转故障 / Config or input anomaly goes to fault
ELSE
CASE _eState OF

    E_DL_CondPotState.eIdle:               // 空闲：使能即进就绪
        IF bEnable THEN
            _eState := E_DL_CondPotState.eReady; // 进就绪 / To ready
        END_IF

    E_DL_CondPotState.eReady:              // 就绪：液位达启位开排
        IF NOT bEnable THEN
            _eState := E_DL_CondPotState.eIdle; // 撤使能回空闲 / Disabled back to idle
        ELSIF _fLevelEff >= fPumpLevelHiPct THEN
            IF uDrainCount < DL_POT_CNT_MAX THEN
                uDrainCount := uDrainCount + 1; // 排放计数递增（饱和不回绕） / Drain counter increment, saturated
            END_IF
            _eState := E_DL_CondPotState.eDraining; // 进排放 / To draining
        END_IF

    E_DL_CondPotState.eDraining:           // 排放中：降至停位关阀或超时判堵
        IF fbDrainMax.Q AND (_fLevelEff > fPumpLevelLoPct) THEN
            _eState := E_DL_CondPotState.eTimeout; // 超时液位未降，判堵塞 / Timeout without level drop, clog
        ELSIF _fLevelEff <= fPumpLevelLoPct THEN
            _eState := E_DL_CondPotState.eReady; // 降至停位，回就绪（阀在段 7 关） / Level at the stop threshold, back to ready
        ELSIF NOT bEnable THEN
            _eState := E_DL_CondPotState.eIdle; // 撤使能回空闲 / Disabled back to idle
        END_IF

    E_DL_CondPotState.eTimeout:            // 排放超时：等复位或液位自行回落
        IF bReset OR (_fLevelEff <= fPumpLevelLoPct) THEN
            _eState := E_DL_CondPotState.eReady; // 解除回就绪 / Cleared back to ready
        END_IF

    E_DL_CondPotState.eFault:              // 故障：复位沿且原因消失回空闲
        IF bReset AND (NOT _bHystBad) THEN
            _eState := E_DL_CondPotState.eIdle; // 回空闲 / Back to idle
        END_IF

    ELSE                                   // 非法状态兜底（R21：CASE 必带 ELSE）
        _bIllegal := TRUE;                 // 标记非法状态 / Flag the illegal state
        _eState   := E_DL_CondPotState.eFault; // 回故障态（阀关） / Back to fault, valve closed
END_CASE
END_IF

(*------------------------------------------------------------------------------
 * 段 7｜输出置位与码位出口（故障/超时态阀显式关——安全侧）
 *      Output assignment and codes, valve explicitly closed on fault
 *-----------------------------------------------------------------------------*)
bDrainOut := (_eState = E_DL_CondPotState.eDraining) AND bEnable AND (NOT _bHystBad); // 仅排放中且合法时开阀 / Valve open only while draining and legal
ePotState := _eState;                       // 相位出口 / Phase outlet

IF _bIllegal THEN
    eErr   := 16#0005_0323;                 // 故障级：状态机兜底 / Fault: state machine fallback
    bError := TRUE;                         // 置故障标志 / Raise the fault flag
ELSIF _bHystBad THEN
    eErr   := 16#0005_0321;                 // 故障级：迟滞倒置或非有限（R90 复用） / Fault: inversion or non-finite, code reused
    bError := TRUE;                         // 置故障标志 / Raise the fault flag
ELSIF _eState = E_DL_CondPotState.eTimeout THEN
    eErr   := 16#0005_0322;                 // 故障级：排放超时判堵塞 / Fault: drain timeout, clog suspected
    bError := TRUE;                         // 置故障标志 / Raise the fault flag
ELSIF _bLevelInfo THEN
    eErr := 16#0005_01E8;                   // 信息级：液位域外已钳位 / Info: level clamped
END_IF

bValid := (NOT bError) AND (_eState <> E_DL_CondPotState.eIdle); // 空闲/故障输出不可用 / Outputs unusable in idle or fault
END_FUNCTION_BLOCK

(* ---- FB_DL_SteamHeaderSplit.st ---- *)
(*
  FB_DL_SteamHeaderSplit  —  蒸汽母管多支路分程分配 / Steam header multi-branch split-range allocation
  分类 Category : DL_Process
  码位 Code     : 16#06_0_93
  版本 Version  : 1.0.0
  溯源 Source   : ModPID 分程控制语义借鉴 · clean-room 实现，仅借分类/参数域/命名，未复制源码
  功能 Function : 1) 母管压力偏差折算总需水率（P 调节口径），按支路优先级顺序分配到各支路阀位输出域；
                  2) 每支路一个 FB_DL_SplitRangeControl 实例承载本支路输出域映射（复用多实例）；
                  3) 逐支路阀位输出钳到本支路行程域。
  边界 Boundary : ① 支路数为 0 拒运行（组态闸）；
                  ② 优先级重复出厂报码（分配顺序不可定即拒算）；
                  ③ 母管压力无效时全支路回安全位（输出域下限）并冻结；
                  ④ 分程区间必须无缝覆盖且不重叠（重叠/空洞出厂报码）；
                  ⑤ 输出三行同向：总需求 → 逐支路阀位 → 分配完成标志。
  依赖 Depends  : FB_DL_SplitRangeControl × 4（逐支路输出域映射，每拍无条件调用）

  码表 Error codes（本件子码步进 16#30 · 本格 93 与既有 9X 子码段冲突，错位至 C3/D3 避让）:
    16#0002_06C3 故障级：组态非法（支路数越界 / 优先级重复 / 分程区间重叠或空洞 / 压力设定 <= 0）
    16#0002_06D3 故障级：相 ID 越界（枚举兜底路径）
    16#0002_06B3 信息级：母管压力无效全支路回安全位冻结（不置 bError）
*)

TYPE E_DL_ShsPhase :
(
    eIdle    := 0,   // 空闲（全支路安全位）/ Idle, all branches at safe position
    eSplit   := 10,  // 分程分配中 / Split allocation running
    eFrozen  := 20,  // 压力无效冻结 / Frozen by invalid header pressure
    eFault   := 90   // 组态故障锁定 / Configuration fault locked
);
END_TYPE

FUNCTION_BLOCK FB_DL_SteamHeaderSplit
VAR_INPUT
    bEnable       : BOOL;                           // 总使能，FALSE 全支路安全位 / Master enable
    bReset        : BOOL;                           // 复位，上升沿清组态故障 / Reset, clears configuration fault
    fHeaderMPa    : REAL;                           // 母管压力实测 [MPa] / Header pressure [MPa]
    fSetMPa       : REAL := 1.0;                    // 母管压力设定 [MPa]，域 > 0 / Header pressure setpoint [MPa]
    fKpPerMPa     : REAL := 100.0;                  // 压力-需求增益 [%/MPa]，域 > 0 / Pressure-to-demand gain [%/MPa]
    nBranchCount  : INT := 3;                       // 支路数 [路]，1..4 / Branch count
    aPriority     : ARRAY[1..4] OF USINT;           // 支路优先级 [1 = 最先分配] / Branch priority, 1 = first
    aDomainLo     : ARRAY[1..4] OF REAL;            // 支路阀位输出域下限 [%] / Branch output domain low [%]
    aDomainHi     : ARRAY[1..4] OF REAL;            // 支路阀位输出域上限 [%] / Branch output domain high [%]
    fSafePosPct   : REAL := 0.0;                    // 安全位阀位 [%] / Safe position [%]
    fEps          : REAL := 1.0E-6;                 // 浮点判零容差 [1] / Floating zero tolerance
END_VAR
VAR_OUTPUT
    afValvePct    : ARRAY[1..4] OF REAL;            // 逐支路分程阀位 [%] / Per-branch split valve position [%]
    bAllocDone    : BOOL;                           // 本拍分配完成标志 / Allocation done this scan
    bFrozen       : BOOL;                           // 压力无效冻结标志 / Frozen by invalid pressure
    bError        : BOOL;                           // 故障标志，与故障级码配对 / Fault flag
    uErrorId      : UDINT;                          // 事件码，0 = 无事件 / Event code
    eStateOut     : E_DL_ShsPhase;                  // 状态机当前态，段尾单点映射 / Phase mapped at tail
END_VAR
VAR
    _eState       : E_DL_ShsPhase := E_DL_ShsPhase.eIdle;  // 内部状态 / Internal state
    afbSplit      : ARRAY[1..4] OF FB_DL_SplitRangeControl;  // 逐支路分程实例（无条件调用）/ Per-branch split-range instance
    rtrReset      : R_TRIG;                         // 复位沿 / Reset edge
    bCfgOk        : BOOL;                           // 组态合法标志 / Configuration valid
    bHdrOk        : BOOL;                           // 母管压力本拍有效 / Header pressure valid
    fDemand       : REAL;                           // 总需求 [%] 0..100 / Total demand [%]
    fRemain       : REAL;                           // 剩余需求 [%] / Remaining demand [%]
    bAllocated    : ARRAY[1..4] OF BOOL;            // 支路已分配掩码 / Branch allocated mask
    afCtrl        : ARRAY[1..4] OF REAL;            // 逐支路需求输入 [%] / Per-branch demand input [%]
    afSpan        : ARRAY[1..4] OF REAL;            // 逐支路域跨度 [%] / Per-branch domain span [%]
    nRank         : USINT;                          // 当前分配序位 / Current allocation rank
    nB            : INT;                            // 支路遍历索引 / Branch loop index
    nFound        : INT;                            // 序位命中支路号 / Branch hit at rank
    uPrioSeen     : ARRAY[1..4] OF USINT;           // 优先级查重表 / Priority duplicate table
    uFault        : UDINT;                          // 锁存故障码 / Latched fault code
    uInfo         : UDINT;                          // 信息级码 / Information code
END_VAR
VAR CONSTANT
    DL_SHS_BMAX   : INT := 4;                       // 支路数上限 [路] / Branch count upper bound
    DL_SHS_INFMAX : REAL := 1.0E30;                 // 压力有限值幅值上限 [MPa] / Pressure finite bound [MPa]
END_VAR

(* === 段 0 · 实例刷新 === *)
rtrReset(CLK := bReset);                          // 每拍刷新复位沿

(* === 段 1 · 组态闸（支路数 / 优先级查重 / 分程区间覆盖性）=== *)
bCfgOk := (nBranchCount >= 1) AND (nBranchCount <= DL_SHS_BMAX)   // 支路数域闸（0 拒运行）
          AND (fSetMPa > fEps) AND (fKpPerMPa > fEps)              // 设定与增益正域
          AND (fSetMPa = fSetMPa) AND (fKpPerMPa = fKpPerMPa);     // NaN 自反
FOR nB := 1 TO DL_SHS_BMAX DO
    uPrioSeen[nB] := 0;                           // 查重表清零
END_FOR
FOR nB := 1 TO nBranchCount DO
    IF (aPriority[nB] >= USINT#1) AND (aPriority[nB] <= USINT#4) THEN
        uPrioSeen[aPriority[nB]] := uPrioSeen[aPriority[nB]] + USINT#1;   // 优先级出现计数（越界优先级按重复计）
    ELSE
        bCfgOk := FALSE;                          // 优先级越域：组态非法
    END_IF
    bCfgOk := bCfgOk AND (aDomainHi[nB] > aDomainLo[nB] + fEps)   // 单支路域不倒置
              AND (aDomainLo[nB] = aDomainLo[nB]) AND (aDomainHi[nB] = aDomainHi[nB]);  // NaN 自反
END_FOR
FOR nB := 1 TO nBranchCount DO
    bCfgOk := bCfgOk AND (uPrioSeen[nB] = USINT#1);   // 每个序位恰好一次（重复/缺位均非法）
END_FOR
FOR nB := 2 TO nBranchCount DO
    bCfgOk := bCfgOk AND (ABS(aDomainLo[nB] - aDomainHi[nB - 1]) < 1.0E-3);  // 相邻域无缝覆盖（容差内贴接）
END_FOR
IF NOT bCfgOk THEN
    uFault := 16#0002_06C3;                       // 故障级：组态非法（含优先级重复与区间重叠/空洞）
END_IF
IF rtrReset.Q AND bCfgOk THEN
    uFault := 16#0000;                            // 复位沿清锁存（解除路径可达）
END_IF
uInfo := 16#0000;                                 // 信息码每拍清零
bHdrOk := (fHeaderMPa = fHeaderMPa) AND (fHeaderMPa >= 0.0) AND (fHeaderMPa < DL_SHS_INFMAX);  // 压力域闸

(* === 段 2 · 总需求折算与按序位残余分配（本拍重算）=== *)
bAllocDone := FALSE;                              // 分配完成本拍重算
fDemand := 0.0;                                   // 需求缺省 0（安全位口径）
FOR nB := 1 TO DL_SHS_BMAX DO
    afCtrl[nB] := 0.0;                            // 支路需求输入清零（安全位口径）
    afSpan[nB] := 0.0;                            // 跨度缺省 0
END_FOR
IF bCfgOk AND bHdrOk AND bEnable THEN
    fDemand := (fSetMPa - fHeaderMPa) * fKpPerMPa;  // 偏差折算需求 [%]（压力低 → 需求大）
    IF fDemand > 100.0 THEN
        fDemand := 100.0;                         // 需求上限钳位
    END_IF
    IF fDemand < 0.0 THEN
        fDemand := 0.0;                           // 需求下限钳位
    END_IF
    fRemain := fDemand;                           // 剩余需求起值
    FOR nRank := 1 TO USINT#4 DO                  // 按优先级序位 1..4 顺序分配（残余递减）
        nFound := 0;                              // 序位命中支路清零
        FOR nB := 1 TO nBranchCount DO
            IF (aPriority[nB] = nRank) AND (nFound = 0) THEN
                nFound := nB;                     // 找到本序位支路
            END_IF
        END_FOR
        bAllocated[nRank] := FALSE;               // 分配掩码先清
        IF nFound > 0 THEN
            bAllocated[nRank] := TRUE;            // 本序位已分配
            afSpan[nFound] := aDomainHi[nFound] - aDomainLo[nFound];   // 本支路域跨度 [%]
            afCtrl[nFound] := fRemain;            // 需求输入 = 当前残余（段 3 内按跨度钳位消化）
            IF fRemain > afSpan[nFound] THEN
                fRemain := fRemain - afSpan[nFound];   // 本支路域已耗尽：残余递减传下序位
            ELSE
                fRemain := 0.0;                   // 残余被本支路消化完
            END_IF
        END_IF
    END_FOR
    bAllocDone := TRUE;                           // 分配完成
ELSIF bCfgOk AND ((NOT bHdrOk) OR (NOT bEnable)) THEN
    uInfo := 16#0002_06B3;                        // 信息级：压力无效/失能全支路安全位冻结
END_IF

(* === 段 3 · 逐支路分程实例（无条件调用）与输出域钳位 === *)
FOR nB := 1 TO DL_SHS_BMAX DO
    afbSplit[nB](bEnable := bCfgOk AND bHdrOk AND bEnable AND bAllocated[nB],   // 本支路参与分配
                 fCtrlIn := afCtrl[nB],             // 本支路需求输入
                 fGap := 0.0,                       // 支路间无中央死区（无缝覆盖组态）
                 rCtrlMax := MAX(afSpan[nB], fEps), // 满量程 = 本支路域跨度（分母防零）
                 rOutHeatMin := aDomainLo[nB],      // 本支路域下限（映射到热通道）
                 rOutHeatMax := aDomainHi[nB],      // 本支路域上限
                 rOutCoolMin := aDomainLo[nB],      // 冷通道复用同域（单通道口径）
                 rOutCoolMax := aDomainHi[nB]);     // 实例每拍无条件调用
    IF bCfgOk AND bHdrOk AND bEnable AND (nB <= nBranchCount) AND afbSplit[nB].bHeatActive THEN
        afValvePct[nB] := afbSplit[nB].fOutHeat;  // 分配中：跟随实例输出
    ELSE
        afValvePct[nB] := fSafePosPct;            // 未参与/冻结/失能：安全位
    END_IF
    IF afValvePct[nB] > aDomainHi[nB] THEN
        afValvePct[nB] := aDomainHi[nB];          // 输出钳到本支路域上限
    END_IF
    IF afValvePct[nB] < aDomainLo[nB] THEN
        afValvePct[nB] := aDomainLo[nB];          // 输出钳到本支路域下限
    END_IF
END_FOR

(* === 段 4 · 主状态机（ENUM + CASE，含 ELSE 兜底）=== *)
CASE _eState OF
E_DL_ShsPhase.eIdle :
    IF uFault <> 16#0000 THEN
        _eState := E_DL_ShsPhase.eFault;          // 故障优先
    ELSIF bEnable AND bCfgOk AND (NOT bHdrOk) THEN
        _eState := E_DL_ShsPhase.eFrozen;         // 压力无效进冻结
    ELSIF bEnable AND bCfgOk AND bHdrOk THEN
        _eState := E_DL_ShsPhase.eSplit;          // 进分程相
    END_IF

E_DL_ShsPhase.eSplit :
    IF (uFault <> 16#0000) OR (NOT bEnable) THEN
        _eState := E_DL_ShsPhase.eFault;          // 故障/失能转出
    ELSIF NOT bHdrOk THEN
        _eState := E_DL_ShsPhase.eFrozen;         // 压力无效转冻结
    END_IF

E_DL_ShsPhase.eFrozen :
    IF bHdrOk AND bEnable AND (uFault = 16#0000) THEN
        _eState := E_DL_ShsPhase.eSplit;          // 压力恢复回分程（解除路径可达）
    END_IF

E_DL_ShsPhase.eFault :
    IF uFault = 16#0000 THEN
        _eState := E_DL_ShsPhase.eIdle;           // 解锁回空闲
    END_IF

ELSE
    _eState := E_DL_ShsPhase.eFault;              // 非法状态拦截
    uFault := 16#0002_06D3;                       // 故障级：相 ID 越界
END_CASE
bFrozen := (_eState = E_DL_ShsPhase.eFrozen) OR (_eState = E_DL_ShsPhase.eFault);  // 冻结标志段尾单点映射

(* === 段 5 · 输出映射 === *)
bError := (uFault <> 16#0000);                    // 故障标志仅由故障级码置位（R45 配对）
IF bError THEN
    uErrorId := uFault;                           // 故障级优先上报
ELSE
    uErrorId := uInfo;                            // 否则上报信息级码
END_IF
eStateOut := _eState;                             // 输出枚举段尾单点映射（N2 规则）
END_FUNCTION_BLOCK

(* ---- FB_DL_SteamTrapDiagTrend.st ---- *)
(*==============================================================================
 * 组件名称 (Component)  : FB_DL_SteamTrapDiagTrend
 * 所属子库 (Sublibrary) : DL_Process
 * 归属目录 (Directory)  : C:\Library\DL_Process
 * 当前版本 (Version)    : 1.0.0
 * 分类/来源标签         : 功能块（FUNCTION_BLOCK）· 过程诊断 · 疏水阀趋势
 *                         industry-pool / steam-system / trend-diagnosis
 * 兼容性   (Platform)   : CODESYS 3.5 / TwinCAT 3 / 汇川 InoProShop / 施耐德
 *                         Machine Expert；仅用 Standard.library 的 TON
 * 溯源声明 (Provenance) : 道莅自研 clean-room——只借公开规范条款与工程惯例，零代码行复制。
 * 功能一句话 (Summary)  : 以过冷度（管线饱和温度与阀前温度之差）为判据，学习窗
 *                         建立基线后监视温差趋势，四级判定蒸汽泄漏等级。
 *
 * 本件存在的意义 (Why this unit exists)：
 *   疏水阀失效开路（直排蒸汽）是蒸汽管网最大的隐性损失。健康阀的过冷度稳定在
 *   基线带内，阀失效后过冷度向零收敛。本件把「过冷度相对基线的收敛程度」变成
 *   四级可观测等级，绝对判据与趋势速率双通道互证，避免单阈值误报。
 *
 * 功能描述 (Function)   : 空闲相等使能转学习；学习相按节拍采样过冷度累加，
 *                         窗满且样本足则建基线（信息级 3000）转监视；窗满样本
 *                         不足回退默认基线并报 3002（保守降级不阻塞监视）；监视
 *                         相按过冷度与基线之比分级（0.7/0.5/0.3），EWMA 趋势以
 *                         K/h 输出。输入非有限冻结评估（3001），非物理跳变冻结
 *                         转重学习（3003）。
 * 与既有件边界 (Boundary): 前置件 FB_DL_SteamTrapMonitor 做单点判定；本件做
 *                         趋势累积与分级，二者正交可级联。
 * 码位说明 (Codes)      : 信息 16#0006_3000 学习完成基线建立
 *                         故障 16#0006_3001 输入非有限，评估冻结
 *                         故障 16#0006_3002 学习窗超时样本不足，基线回退默认
 *                         故障 16#0006_3003 非物理跳变，判定冻结转重学习
 *                         段 16#06_0_00~04 首槽信息级、次槽起故障级。
 * 依赖说明 (Depends)    : 无 DL_ 内部依赖；仅 Standard.library 的 TON。
 * 红线自检 (Redline)    : 零全局依赖 ｜ 零 VAR_EXTERNAL ｜ 零 %I/%Q ｜ 纯 IEC 标准库
 *                         浮点比较全部带 fEps 容差 ｜ NaN/Inf 精确判据拦截
 *                         ENUM 配 CASE 且 ELSE 兜底 ｜ 定时器每周期无条件刷新
 *                         全变量双语同行注释 ｜ 故障锁存回放且有可达解除路径
 * 修订历史 (Revision)   : 2026-11-18  v1.0.0  首版入库（R32 · 批 2）
 *============================================================================*)

FUNCTION_BLOCK FB_DL_SteamTrapDiagTrend
VAR_INPUT
    bRun          : BOOL;                   // 诊断使能，假则回空闲并清判定 / Enable, FALSE returns to idle
    fTrapTempC    : LREAL;                  // 阀前温度 [degC] / Trap body temperature
    fLineTempC    : LREAL;                  // 管线饱和温度基准 [degC] / Line saturation reference temperature
    fDTBaseDef    : LREAL := 15.0;          // 默认基线过冷度 [K]，学习失败回退值 / Default baseline subcooling
    fRatioWatch   : LREAL := 0.7;           // 关注级阈值 [比值]，低于此进入关注 / Watch level ratio threshold
    fRatioSuspect : LREAL := 0.5;           // 可疑级阈值 [比值] / Suspect level ratio threshold
    fRatioLeak    : LREAL := 0.3;           // 泄漏级阈值 [比值] / Leak level ratio threshold
    fEps          : LREAL := 1.0E-6;        // 浮点判零容差 [实数域] / Floating zero tolerance
    tLearnWin     : TIME  := T#30M;         // 学习窗时长 [s] / Learning window duration
    tSample       : TIME  := T#10S;         // 采样节拍 [s] / Sampling pace period
END_VAR
VAR_OUTPUT
    eLevel    : (eLevelOk := 0, eLevelWatch := 1, eLevelSuspect := 2, eLevelLeak := 3);  // 泄漏等级枚举 / Leak level enum
    fBaseDT   : LREAL;                  // 已建立基线过冷度 [K] / Established baseline subcooling
    fDTNow    : LREAL;                  // 当前过冷度 [K] / Current subcooling
    fTrendKpH : LREAL;                  // 过冷度趋势 [K/h]，负值为向零收敛 / Subcooling trend, negative converges to zero
    bDiag     : BOOL;                   // 判定有效标志，监视相且数据有效为真 / TRUE when the verdict is valid
    bError    : BOOL;                   // 故障标志，与故障码配对 / Fault flag paired with codes
    uErrorId  : UDINT;                  // 事件码，0 表示无事件 / Event code, zero means none
END_VAR
VAR
    eState    : (eIdle := 0, eLearning := 1, eMonitor := 2);    // 状态机：空闲/学习/监视 / State machine
    tonLearn  : TON;    // 学习窗定时器 [s]，每拍无条件刷新 / Learning window timer
    tonPace   : TON;    // 采样节拍定时器 [s]，每拍无条件刷新 / Sampling pace timer
    bSigOk    : BOOL;   // 输入有效标志 / Input validity flag
    fSumDT    : LREAL;  // 学习相过冷度累加和 [K] / Learning-phase subcooling sum
    nSamples  : UDINT;  // 有效样本数 [个] / Valid sample count
    fDTLast   : LREAL;  // 上拍过冷度快照 [K] / Previous subcooling snapshot
    bHavePrev : BOOL;   // 快照有效标志 / Snapshot availability flag
    fTrendEw  : LREAL;  // 趋势 EWMA 内部值 [K/h] / Trend EWMA internal value
    fPaceS    : LREAL;  // 采样节拍秒值 [s]，由 tSample 一次性导出 / Pace in seconds, derived once
    uCodeLatch: UDINT;  // 故障锁存码 [码]，故障相回放 / Latched fault code
    uInfoCode : UDINT;  // 信息级单拍码 [码]，出口装配后即清 / One-shot info code, cleared after assembly
END_VAR
VAR CONSTANT
    DL_STT_MINSAMP : INT   := 10;       // 学习窗最小样本数 [个] / Minimum learning samples
    DL_STT_JUMP    : LREAL := 50.0;     // 单拍非物理跳变门限 [K] / Non-physical jump limit
    DL_STT_TAU     : LREAL := 0.1;      // 趋势 EWMA 平滑系数 [比值] / Trend EWMA smoothing factor
    DL_STT_H2S     : LREAL := 3600.0;   // 每小时秒数 [s/h] / Seconds per hour
    DL_STT_MS2S    : LREAL := 1000.0;   // 毫秒到秒系数 [ms/s] / Milliseconds per second
END_VAR

(* 段 1｜定时器无条件周期刷新（红线 7）：两实例每拍先触发 / Timers refreshed unconditionally every scan *)
tonLearn(IN := (eState = eLearning) AND bRun, PT := tLearnWin);     // 学习窗计时 / Learning window timing
tonPace(IN := bRun, PT := tSample);                                 // 采样节拍计时 / Sampling pace timing
IF fPaceS < 0.0001 THEN
    fPaceS := DINT_TO_LREAL(TIME_TO_DINT(tSample)) / DL_STT_MS2S;   // 节拍秒值一次导出 / Derive pace seconds once
END_IF

(* 段 2｜当前过冷度与输入有效性（每拍计算，判据门控挂状态量）/ Current subcooling and validity each scan *)
fDTNow := fLineTempC - fTrapTempC;                                  // 过冷度导出 / Derive subcooling
bSigOk := (fTrapTempC = fTrapTempC) AND (fLineTempC = fLineTempC)   // NaN 自反判据 / NaN reflexivity
          AND (ABS(fTrapTempC) < 1.0E308) AND (ABS(fLineTempC) < 1.0E308)   // Inf 上限判据 / Inf limit
          AND (fDTNow >= -fEps);                                    // 过冷度非负物理约束 / Non-negativity

(* 段 3｜状态机主分派（ENUM 配 CASE，ELSE 兜底）/ State dispatch with ELSE interception *)
CASE eState OF

    eIdle:
        bDiag := FALSE;                 // 空闲不出判定 / No verdict in idle
        eLevel := eLevelOk;             // 默认级 / Default level
        fSumDT := 0.0;                  // 清累加 / Clear the sum
        nSamples := 0;                  // 清计数 / Clear the count
        fTrendEw := 0.0;                // 清趋势 / Clear the trend
        bHavePrev := FALSE;             // 清快照 / Clear the snapshot
        IF bRun AND bSigOk THEN
            eState := eLearning;        // 拍 N 空闲相满足条件，拍 N+1 进入学习 / Idle to learning next scan
        END_IF

    eLearning:
        (* 本拍行为：节拍到点且数据有效则采样累加；退出条件 = 窗满 AND 样本足（双条件）
         * This scan: sample on pace tick; exit needs window done AND enough samples *)
        IF NOT bSigOk THEN
            uCodeLatch := 16#0006_3001; // 故障：输入非有限 / Fault: non-finite input
        ELSIF tonPace.Q THEN
            fSumDT := fSumDT + fDTNow;  // 累加 / Accumulate
            nSamples := nSamples + 1;   // 计数 / Count
        END_IF
        IF tonLearn.Q AND (nSamples >= INT_TO_UDINT(DL_STT_MINSAMP)) THEN
            fBaseDT := fSumDT / UDINT_TO_LREAL(nSamples);   // 均值基线 / Mean baseline
            uCodeLatch := 16#0000_0000;                     // 学习成功清除锁存 / Success clears the latch
            uInfoCode := 16#0006_3000;                      // 信息级：基线建立（单拍）/ Info: baseline built, one shot
            eState := eMonitor;                             // 拍 N+1 转监视 / To monitor next scan
        ELSIF tonLearn.Q AND (nSamples < INT_TO_UDINT(DL_STT_MINSAMP)) THEN
            fBaseDT := fDTBaseDef;      // 保守回退默认基线，不阻塞监视 / Conservative fallback, monitoring unblocked
            uCodeLatch := 16#0006_3002; // 故障：样本不足已回退 / Fault: insufficient samples, fallback
            eState := eMonitor;         // 拍 N+1 转监视 / To monitor next scan
        END_IF

    eMonitor:
        bDiag := bSigOk;                // 判定有效随数据有效 / Verdict valid with the data
        IF NOT bSigOk THEN
            uCodeLatch := 16#0006_3001; // 故障：输入非有限，判定冻结 / Fault: non-finite, frozen
        ELSIF ABS(fBaseDT) < fEps THEN
            uCodeLatch := 16#0006_3003; // 故障：基线异常，转重学习 / Fault: bad baseline, relearn
            fSumDT := 0.0;              // 清累加 / Clear the sum
            nSamples := 0;              // 清计数 / Clear the count
            eState := eLearning;        // 拍 N+1 转学习 / To learning next scan
        ELSE
            (* 非物理跳变闸：单拍变化超限说明传感器异常，冻结并重学习 / Jump gate: freeze and relearn *)
            IF bHavePrev AND (ABS(fDTNow - fDTLast) > DL_STT_JUMP) THEN
                uCodeLatch := 16#0006_3003;     // 故障：非物理跳变 / Fault: non-physical jump
                fSumDT := 0.0;                  // 清累加 / Clear the sum
                nSamples := 0;                  // 清计数 / Clear the count
                eState := eLearning;            // 拍 N+1 转学习 / To learning next scan
            ELSE
                (* 分级判据：过冷度相对基线的收敛程度 / Grading: convergence relative to the baseline *)
                IF fDTNow < (fRatioLeak * fBaseDT) THEN
                    eLevel := eLevelLeak;       // 泄漏级 / Leak level
                ELSIF fDTNow < (fRatioSuspect * fBaseDT) THEN
                    eLevel := eLevelSuspect;    // 可疑级 / Suspect level
                ELSIF fDTNow < (fRatioWatch * fBaseDT) THEN
                    eLevel := eLevelWatch;      // 关注级 / Watch level
                ELSE
                    eLevel := eLevelOk;         // 健康级 / Healthy level
                END_IF
                (* 趋势采样：节拍到点且快照有效则算瞬时趋势并 EWMA / Trend sample on pace tick *)
                IF tonPace.Q AND bHavePrev AND (fPaceS > fEps) THEN
                    fTrendEw := fTrendEw * (1.0 - DL_STT_TAU)
                                + ((fDTNow - fDTLast) / fPaceS * DL_STT_H2S) * DL_STT_TAU;  // K/h 瞬时趋势入 EWMA / K/h trend into EWMA
                END_IF
            END_IF
        END_IF

ELSE
    eState := eIdle;                    // 非法状态拦截回空闲 / Illegal state intercepted to idle
    uCodeLatch := 16#0006_3001;         // 故障：状态越界 / Fault: state out of range
END_CASE

(* 段 4｜快照与出口装配 / Snapshot and exit assembly *)
fDTLast := fDTNow;                      // 更新快照供下拍跳变判据 / Update the snapshot for the next scan
bHavePrev := bSigOk;                    // 快照有效随数据有效 / Snapshot valid with the data
fTrendKpH := fTrendEw;                  // 趋势输出 / Trend output
IF NOT bRun THEN
    uCodeLatch := 16#0000_0000;         // 撤使能清故障（可达解除路径）/ Run drop clears faults, reachable reset
END_IF
bError   := (uCodeLatch <> 16#0000_0000);   // 故障锁存回放 / Latched fault replay
IF uCodeLatch <> 16#0000_0000 THEN
    uErrorId := uCodeLatch;             // 故障码优先回放 / Fault code replayed first
    uInfoCode := 16#0000_0000;          // 故障压过信息码 / Fault overrides the info code
ELSE
    uErrorId := uInfoCode;              // 无故障时放信息码 / Info code when no fault
    uInfoCode := 16#0000_0000;          // 信息码单拍清零 / Info code cleared next scan
END_IF
END_FUNCTION_BLOCK

(* ---- FB_DL_StratificationGuard.st ---- *)
(*
  FB_DL_StratificationGuard  —  水箱温度分层监视与混温抑制 / Tank thermal stratification monitor with mixing suppression
  分类 Category : DL_Process
  码位 Code     : 16#06_0_88
  版本 Version  : 1.0.0
  溯源 Source   : Modular PID 语义借鉴 · clean-room 实现，仅借分类/参数域/命名，未复制源码
  功能 Function : 1) 上下点温差带迟滞判据（起动门限 > 停止门限），防混水泵频繁启停；
                  2) 两点任一无效时冻结判定并保持上次输出；
                  3) 混温请求与主机启动命令互斥仲裁，同拍双真取安全侧（抑制混温、让主机优先）。
  边界 Boundary : ① 温差判据带迟滞（fDiffOnC 必须 > fDiffOffC，否则组态报码）；
                  ② 两点任一无效时冻结判定并保持上次输出（bFreeze）；
                  ③ 混温请求与主机启动命令互斥仲裁，同拍双真取安全侧；
                  ④ 仲裁态三行同向：混温请求 → 温差记录 → 冻结标志。
  依赖 Depends  : None

  码表 Error codes（本件子码步进 16#10，避让邻件码位）:
    16#0002_0688 故障级：迟滞门限非法（fDiffOnC <= fDiffOffC 或门限 <= 0）
    16#0002_0698 故障级：相 ID 越界（枚举兜底路径）
    16#0002_06A8 信息级：仲裁互斥生效（主机启动优先，混温请求被抑制，不置 bError）
*)

TYPE E_DL_StratPhase :
(
    eIdle    := 0,   // 空闲 / Idle
    eMonitor := 10,  // 温差监视 / Differential monitoring
    eMixOn   := 20,  // 混温运行 / Mixing active
    eFreeze  := 30,  // 无效点冻结 / Frozen by invalid points
    eFault   := 90   // 故障锁定 / Fault locked
);
END_TYPE

FUNCTION_BLOCK FB_DL_StratificationGuard
VAR_INPUT
    bEnable      : BOOL;                          // 总使能，FALSE 回空闲停泵 / Master enable
    bReset       : BOOL;                          // 复位，上升沿清故障 / Reset, clears fault
    fTempTopC    : REAL;                          // 水箱上部温度 [degC]，域 −20~120 / Upper tank temperature [degC]
    bTopValid    : BOOL := TRUE;                  // 上部温度通道有效 / Upper channel valid
    fTempBotC    : REAL;                          // 水箱下部温度 [degC]，域 −20~120 / Lower tank temperature [degC]
    bBotValid    : BOOL := TRUE;                  // 下部温度通道有效 / Lower channel valid
    fDiffOnC     : REAL := 5.0;                   // 混温起动温差门限 [degC]，域 > 0 / Mixing start threshold [degC]
    fDiffOffC    : REAL := 2.0;                   // 混温停止温差门限 [degC]，域 > 0 且 < 起动门限 / Mixing stop threshold
    fDiffMaxC    : REAL := 30.0;                  // 温差物理域上限 [degC]，超此值判传感器异常 / Differential domain high
    bHostStartCmd: BOOL;                          // 主机启动命令（互斥仲裁输入）/ Host start command for arbitration
    fEps         : REAL := 1.0E-6;                // 浮点判零容差 [1] / Floating zero tolerance
END_VAR
VAR_OUTPUT
    fDiffC       : REAL;                          // 上下点温差 [degC]（上 − 下）/ Top-minus-bottom differential [degC]
    bMixPumpReq  : BOOL;                          // 混温泵请求 [开关] / Mixing pump request
    bFreeze      : BOOL;                          // 判定冻结标志（保持型）/ Judgment frozen, held
    bArbitActive : BOOL;                          // 仲裁互斥生效标志 / Arbitration active flag
    bError       : BOOL;                          // 故障标志，与故障级码配对 / Fault flag paired with fault codes
    uErrorId     : UDINT;                         // 事件码，0 = 无事件 / Event code, 0 = none
    eStateOut    : E_DL_StratPhase;               // 状态机当前态，段尾单点映射 / Phase mapped at tail
END_VAR
VAR
    _eState      : E_DL_StratPhase := E_DL_StratPhase.eIdle;  // 内部状态 / Internal state
    rtrReset     : R_TRIG;                        // 复位沿 / Reset edge
    bPtsOk       : BOOL;                          // 两点均有效 / Both points valid
    bCfgOk       : BOOL;                          // 门限组态合法 / Thresholds valid
    bMixLatched  : BOOL;                          // 混温请求锁存（迟滞用）/ Mixing request latch for hysteresis
    fDiffBuf     : REAL;                          // 本拍温差 [degC] / Differential this scan
    uFault       : UDINT;                         // 锁存故障码 / Latched fault code
    uInfo        : UDINT;                         // 信息级码 / Information code
END_VAR
VAR CONSTANT
    DL_STR_TMIN  : REAL := -20.0;                 // 温度物理域下限 [degC] / Temperature domain low
    DL_STR_TMAX  : REAL := 120.0;                 // 温度物理域上限 [degC] / Temperature domain high
END_VAR

(* === 段 0 · 实例刷新（无条件周期调用）=== *)
rtrReset(CLK := bReset);                          // 每拍刷新复位沿

(* === 段 1 · 组态闸与测点域闸 === *)
bCfgOk := (fDiffOnC > fEps) AND (fDiffOffC > fEps) AND (fDiffOnC > fDiffOffC + fEps)
          AND (fDiffMaxC > fDiffOnC) AND (fDiffOnC = fDiffOnC) AND (fDiffOffC = fDiffOffC);   // 含 NaN 自反
IF NOT bCfgOk THEN
    uFault := 16#0002_0688;                       // 故障级：迟滞门限非法（倒置或非正）
END_IF
IF rtrReset.Q AND bCfgOk THEN
    uFault := 16#0000;                            // 复位沿清锁存（复位路径可达）
END_IF
bPtsOk := bTopValid AND bBotValid
          AND (fTempTopC = fTempTopC) AND (fTempBotC = fTempBotC)          // NaN 自反判据
          AND (ABS(fTempTopC) < 1.0E30) AND (ABS(fTempBotC) < 1.0E30)      // Inf 上限兜底
          AND (fTempTopC >= DL_STR_TMIN) AND (fTempTopC <= DL_STR_TMAX)     // 上点物理域
          AND (fTempBotC >= DL_STR_TMIN) AND (fTempBotC <= DL_STR_TMAX);    // 下点物理域
IF bPtsOk THEN
    fDiffBuf := fTempTopC - fTempBotC;            // 温差 = 上 − 下（正 = 上部更热，分层成立）
ELSE
    fDiffBuf := fDiffC;                           // 无效点：温差保持上次值，不参与判定
END_IF
IF ABS(fDiffBuf) > fDiffMaxC THEN
    uInfo := 16#0002_06A8;                        // 信息级：温差超物理域，疑似传感器异常
    bPtsOk := FALSE;                              // 超域按无效处理，冻结判定
END_IF
fDiffC := fDiffBuf;                               // 温差输出

(* === 段 2 · 主状态机（ENUM + CASE，含 ELSE 兜底）=== *)
CASE _eState OF
E_DL_StratPhase.eIdle :
    bMixPumpReq := FALSE;                         // 空闲停泵
    bFreeze := FALSE;                             // 冻结标志复位
    bMixLatched := FALSE;                         // 迟滞锁存复位
    uInfo := 16#0000;                             // 信息码清零（本拍异常会重新置位）
    IF uFault <> 16#0000 THEN
        _eState := E_DL_StratPhase.eFault;        // 故障优先
    ELSIF bEnable AND (NOT bPtsOk) THEN
        bFreeze := TRUE;                          // 上电即无效：直接冻结
        _eState := E_DL_StratPhase.eFreeze;
    ELSIF bEnable THEN
        _eState := E_DL_StratPhase.eMonitor;      // 进入监视相
    END_IF

E_DL_StratPhase.eMonitor :
    IF NOT bPtsOk THEN
        bFreeze := TRUE;                          // 任一测点无效：冻结判定
        _eState := E_DL_StratPhase.eFreeze;
    ELSE
        bFreeze := FALSE;                         // 两点有效：解冻
        IF (NOT bMixLatched) AND (fDiffC >= fDiffOnC) THEN
            bMixLatched := TRUE;                  // 越起动门限：置请求锁存
            bMixPumpReq := TRUE;                  // 混温请求输出
            _eState := E_DL_StratPhase.eMixOn;
        END_IF
    END_IF

E_DL_StratPhase.eMixOn :
    bMixPumpReq := TRUE;                          // 混温运行
    IF NOT bPtsOk THEN
        bFreeze := TRUE;                          // 测点无效：冻结（请求保持上次值）
        _eState := E_DL_StratPhase.eFreeze;
    ELSIF fDiffC <= fDiffOffC THEN
        bMixLatched := FALSE;                     // 降到停止门限以下：解除（迟滞回差生效）
        bMixPumpReq := FALSE;                     // 停泵
        _eState := E_DL_StratPhase.eMonitor;
    END_IF

E_DL_StratPhase.eFreeze :
    bFreeze := TRUE;                              // 冻结标志保持
    IF bPtsOk THEN
        bFreeze := FALSE;                         // 两点恢复有效：解冻（可到达的解除路径）
        uInfo := 16#0000;                         // 信息码清除
        _eState := E_DL_StratPhase.eMonitor;
    END_IF

E_DL_StratPhase.eFault :
    bMixPumpReq := FALSE;                         // 故障态停泵（安全侧）
    bFreeze := TRUE;                              // 冻结判定
    bMixLatched := FALSE;                         // 迟滞锁存复位
    IF uFault = 16#0000 THEN
        _eState := E_DL_StratPhase.eIdle;         // 解锁回空闲
    END_IF

ELSE
    _eState := E_DL_StratPhase.eFault;            // 非法状态拦截
    uFault := 16#0002_0698;                       // 故障级：相 ID 越界（枚举兜底路径）
    bMixPumpReq := FALSE;                         // 安全侧停泵
END_CASE

(* === 段 3 · 互斥仲裁：混温请求 vs 主机启动命令（同拍双真取安全侧）=== *)
bArbitActive := FALSE;                            // 仲裁标志每拍重算
IF bHostStartCmd AND bMixPumpReq THEN
    bMixPumpReq := FALSE;                         // 安全侧：主机启动优先，抑制混温
    bMixLatched := FALSE;                         // 迟滞锁存同步复位，防下一拍立即复启
    bArbitActive := TRUE;                         // 仲裁互斥生效
    uInfo := 16#0002_06A8;                        // 信息级：仲裁互斥（不置 bError）
END_IF

(* === 段 4 · 输出映射（三行同向：请求 → 温差 → 冻结标志）=== *)
IF NOT bEnable THEN
    bMixPumpReq := FALSE;                         // 失能最高优先停泵
    bArbitActive := FALSE;                        // 失能不算仲裁
END_IF
bError := (uFault <> 16#0000);                    // 故障标志仅由故障级码置位（R45 配对）
IF bError THEN
    uErrorId := uFault;                           // 故障级优先上报
ELSE
    uErrorId := uInfo;                            // 否则上报信息级码
END_IF
eStateOut := _eState;                             // 输出枚举段尾单点映射（N2 规则）
END_FUNCTION_BLOCK

(* ---- FB_DL_StringBarcodeTrace.st ---- *)
// =====================================================================
// FB_DL_StringBarcodeTrace.st
// 电池串条码绑定与工位路由（校验→拼接追溯键→查重→首绑定为准）
// Barcode binding and station routing FB
// 码位: 16#0005_0453 ~ 16#0005_0457 (本件独占 5 槽)
// 修改记录: R29 初版 (按 DISPATCH_R29 序 17)
// =====================================================================
FUNCTION_BLOCK FB_DL_StringBarcodeTrace
VAR_INPUT
    bEnable      : BOOL  := FALSE;    // 使能 / Enable
    bReset       : BOOL  := FALSE;    // 复位（含清重码计数）/ Reset
    bCodeValid   : BOOL  := FALSE;    // 扫码完成有效（脉冲）/ Code valid pulse
    sCode        : STRING(32) := '';  // 扫码内容，32 字符上限 / Scanned code
    sLotKey      : STRING(16) := '';  // 批次键（外部下发）/ Lot key
    uStationIdx  : USINT  := 1;       // 当前工位号 1~99 / Station index
    uStationCnt  : USINT  := 8;       // 工位总数 1~99 / Station count
    uLenMin      : USINT  := 8;       // 码最小长度 1~32 / Min length
    uLenMax      : USINT  := 24;      // 码最大长度 1~32 / Max length
    uDupMax      : USINT  := 3;       // 连续重码报警次数 1~20 / Duplicate alarm count
END_VAR
VAR_OUTPUT
    sBindingKey  : STRING(64);        // 追溯键 Lot|Station|Code / Binding key
    uRouteIdx    : USINT;             // 路由工位号 / Route index
    bRouteValid  : BOOL;              // 路由有效（可放行）/ Route valid
    bDuplicate   : BOOL;              // 重码（首绑定未被覆盖）/ Duplicate
    uDupCnt      : USINT;             // 连续重码计数 / Consecutive duplicate count
    eErr         : UDINT;             // 错误码 / Error code
END_VAR
VAR
    rtrigValid   : R_TRIG;            // 扫码有效沿检测（无条件刷新）/ Code valid edge detector
    aDupCode     : ARRAY[0..31] OF STRING(32);    // 重码环形记录表 / Duplicate ring records
    uDupHead     : USINT;             // 环形写指针 / Ring write pointer
    uDupFill     : USINT;             // 环形已存条数 / Ring filled count
    uIdx         : USINT;             // 查重循环下标 / Search loop index
    uLen         : USINT;             // 码长度 / Code length
    uChar        : USINT;             // 字符循环下标 / Char loop index
    sChar        : STRING(1);         // 单字符临时 / Single char temp
    bCharOK      : BOOL;              // 字符合法标记 / Char valid flag
    uLotLen      : USINT;             // 批次键长度 / Lot key length
    uStLen       : USINT;             // 工位号字符串长度 / Station string length
    uTotalLen    : USINT;             // 拼接结果总长（先算后拼）/ Total result length
    sStTmp       : STRING(8);         // 工位号字符串临时 / Station string temp
    bDupFound    : BOOL;              // 重码命中标记 / Duplicate found flag
    bLockLatch   : BOOL := FALSE;     // 连续重码故障锁存 / Consecutive dup fault latch
    xFirstScan   : BOOL  := TRUE;     // 首扫标记 / First-scan flag
END_VAR

// ---------------------------------------------------------------------
// 代码位表（本件独占，勿复用）:
//   16#0005_0453 信息 绑定成功、码唯一
//   16#0005_0454 故障 sLotKey 为空 / bCodeValid 时 sCode 为空串
//   16#0005_0455 故障 uStationIdx > uStationCnt / uStationCnt = 0 / uLenMin > uLenMax（组态错）
//   16#0005_0456 信息 码格式非法（长度/字符集不符）→ 拒收，bRouteValid=FALSE；拼接超限截断同登记
//   16#0005_0457 故障 bDuplicate 连续 uDupMax 次 → 锁存（uDupCnt ≥ uDupMax）
// ---------------------------------------------------------------------

// ---- 扫码沿检测（无条件刷新，R47 边沿纪律）/ Code valid edge, unconditional ----
rtrigValid(CLK := bCodeValid);  // 沿检测 / Edge detection

// ---- 组态错闸 / Configuration fault gate ----
IF (uStationCnt = 0) OR (uStationIdx > uStationCnt) OR (uLenMin > uLenMax)
   OR (uLenMin = 0) OR (uDupMax = 0) THEN
    bRouteValid := FALSE;       // 路由撤销 / Route invalid
    eErr := 16#0005_0455;       // 故障码 / Fault code
    RETURN;                     // 本拍结束 / End of cycle
END_IF

// ---- 首扫初始化（R16 首扫纪律）/ First-scan initialization ----
IF xFirstScan THEN
    bRouteValid := FALSE;       // 路由初始无效 / Route init invalid
    uRouteIdx := 0;             // 路由号清零 / Route cleared
    xFirstScan := FALSE;        // 清标记 / Clear flag
END_IF

// ---- 复位：清重码计数与重码表 / Reset: clear dup count and table ----
IF bReset THEN
    uDupCnt := 0;               // 计数清零 / Count cleared
    bDuplicate := FALSE;        // 重码复位 / Duplicate reset
    bLockLatch := FALSE;        // 锁存解除 / Latch released
    FOR uIdx := 0 TO 31 DO
        aDupCode[uIdx] := '';   // 重码表清空 / Table cleared
    END_FOR
    uDupHead := 0;              // 指针归零 / Pointer reset
    uDupFill := 0;              // 填充数清零 / Fill reset
END_IF

// ---- 使能撤销 / Disable ----
IF NOT bEnable THEN
    bRouteValid := FALSE;       // 路由撤销 / Route invalid
    bDuplicate := FALSE;        // 重码复位 / Duplicate reset
    eErr := 16#0005_0453;       // 信息级：空闲 / Info: idle
    RETURN;                     // 本拍结束 / End of cycle
END_IF

// ---- 连续重码锁存路径 / Consecutive duplicate latch path ----
IF bLockLatch THEN
    bRouteValid := FALSE;       // 放行撤销 / Route invalid
    eErr := 16#0005_0457;       // 故障码回放 / Fault code replay
    RETURN;                     // 本拍结束 / End of cycle
END_IF

// ---- 非沿拍维持原状 / Non-edge cycles hold state ----
IF NOT rtrigValid.Q THEN
    RETURN;                     // 绑定结果与路由保持 / Binding and route hold
END_IF

// ---- 批次键/码空闸（故障级）/ Empty lot or code gate ----
uLotLen := LEN(sLotKey);        // 批次键长度 / Lot length
uLen := LEN(sCode);             // 码长度 / Code length
IF (uLotLen = 0) OR (uLen = 0) THEN
    bRouteValid := FALSE;       // 路由撤销 / Route invalid
    eErr := 16#0005_0454;       // 故障码 / Fault code
    RETURN;                     // 本拍结束 / End of cycle
END_IF

// ---- 长度校验（越界拒收信息级）/ Length validation ----
IF (uLen < uLenMin) OR (uLen > uLenMax) THEN
    bRouteValid := FALSE;       // 拒收 / Rejected
    eErr := 16#0005_0456;       // 信息级：格式非法 / Info: format invalid
    RETURN;                     // 本拍结束 / End of cycle
END_IF

// ---- 字符集校验：只允许数字与字母 / Charset validation: digits and letters only ----
bCharOK := TRUE;                // 先假设合法 / Assume valid
FOR uChar := 1 TO uLen DO
    sChar := MID(sCode, 1, uChar);      // 取单字符 / Extract char
    // 字典序判数字/大写/小写（纯 IEC 61131-3 字符串比较，不用非标准 ASCII 函数）
    // Lexicographic alnum check, pure IEC string comparison
    IF NOT (((sChar >= '0') AND (sChar <= '9'))
        OR ((sChar >= 'A') AND (sChar <= 'Z'))
        OR ((sChar >= 'a') AND (sChar <= 'z'))) THEN
        bCharOK := FALSE;       // 非数字字母 / Not alnum
    END_IF
END_FOR
IF NOT bCharOK THEN
    bRouteValid := FALSE;       // 拒收 / Rejected
    eErr := 16#0005_0456;       // 信息级：格式非法 / Info: format invalid
    RETURN;                     // uRouteIdx 不变 / Route holds
END_IF

// ---- 查重：环形表线性比对 / Duplicate search in ring table ----
bDupFound := FALSE;             // 命中复位 / Reset hit
FOR uIdx := 0 TO 31 DO
    IF (uIdx < uDupFill) AND (aDupCode[uIdx] = sCode) THEN
        bDupFound := TRUE;      // 命中 / Hit
    END_IF
END_FOR

IF bDupFound THEN
    // 重码：不覆盖首绑定，计数递增 / Duplicate: first binding kept, count up
    bDuplicate := TRUE;         // 重码标志 / Duplicate flag
    uDupCnt := uDupCnt + 1;     // 计数 / Count
    bRouteValid := FALSE;       // 本次不放行 / Not released
    IF uDupCnt >= uDupMax THEN
        bLockLatch := TRUE;     // 连续重码 → 锁存 / Latch on consecutive dups
        eErr := 16#0005_0457;   // 故障码 / Fault code
    ELSE
        eErr := 16#0005_0456;   // 信息级：重码拒收 / Info: duplicate rejected
    END_IF
    RETURN;                     // sBindingKey 保持首次值 / Binding key holds first value
END_IF

// ---- 拼接追溯键：先算后拼（上限 64，超限截 63 并置槽 4）/ Build key: compute length first ----
uStLen := 2;                    // 工位号最多两位数（1~99）/ Station digits max 2
uTotalLen := uLotLen + 1 + uStLen + 1 + uLen;   // Lot + | + St + | + Code / Total length
IF uTotalLen > 64 THEN
    // 超限：截 63 写入并登记（禁越界写）/ Over limit: truncate to 63
    sBindingKey := CONCAT(sLotKey, '|');
    sBindingKey := CONCAT(sBindingKey, USINT_TO_STRING(uStationIdx));
    sBindingKey := CONCAT(sBindingKey, '|');
    sBindingKey := CONCAT(sBindingKey, LEFT(sCode, 63 - uLotLen - 1 - uStLen - 1));   // 截断码 / Truncated code
    bRouteValid := FALSE;       // 键不完整不放行 / Incomplete key, no release
    eErr := 16#0005_0456;       // 信息级：超限截断 / Info: truncated
    RETURN;                     // 本拍结束 / End of cycle
END_IF

sBindingKey := CONCAT(sLotKey, '|');                    // Lot| / Lot|
sBindingKey := CONCAT(sBindingKey, USINT_TO_STRING(uStationIdx));   // +Station / +Station
sBindingKey := CONCAT(sBindingKey, '|');                // +| / +|
sBindingKey := CONCAT(sBindingKey, sCode);              // +Code / +Code

// ---- 首次绑定登记：入环形表（满覆盖最旧并置信息）/ First binding: register into ring ----
aDupCode[uDupHead] := sCode;    // 登记码 / Register code
uDupHead := uDupHead + 1;       // 指针前移 / Pointer advance
IF uDupHead > 31 THEN
    uDupHead := 0;              // 回绕 / Wrap
END_IF
IF uDupFill < 32 THEN
    uDupFill := uDupFill + 1;   // 填充 / Fill
ELSE
    // 表满覆盖最旧：信息级提示（不影响放行逻辑）/ Table full: overwrite oldest
    eErr := 16#0005_0456;       // 信息级 / Info
END_IF

// ---- 绑定成功 / Binding success ----
bDuplicate := FALSE;            // 重码复位 / Duplicate reset
uRouteIdx := uStationIdx;       // 路由号 = 当前工位 / Route = station
bRouteValid := TRUE;            // 放行 / Released
IF eErr <> 16#0005_0456 THEN
    eErr := 16#0005_0453;       // 信息级：绑定成功 / Info: bound
END_IF

END_FUNCTION_BLOCK
